                               //Extractor Cnv FROM CNV1
                           ELSIF (#Destination_Location.Device_Type = 12 AND #Source_Location.Device_Type = 10 AND
                               NOT "Control_DB".ECnv_Sys[#Id].Cnv_Occupied AND
                               "Control_DB".LCnv_Sys[#Id].Cnv_Level[#Destination_Location.Level].Cnv1.Cnv_Occupied)
                           THEN //FROM ECONVEYOR TO CNV1 OR CNV2
                               "Control_DB".ECnv_Sys[#Id].Instruction.Task_ID := INT_TO_UINT("Control_DB".WCS_OPC_Control[#Id].Task_ID);
                               "Control_DB".ECnv_Sys[#Id].Instruction.Task_Metadata := "Control_DB".WCS_OPC_Control[#Id].Task_Metadata;
                               "Control_DB".ECnv_Sys[#Id].Current_Task_Type := INT_TO_UINT("Control_DB".WCS_OPC_Control[#Id].Task_Type);
                               "Control_DB".ECnv_Sys[#Id].Instruction.Transfer_From_ID := "Control_DB".WCS_OPC_Control[#Id].Source_Location;
                               "Control_DB".ECnv_Sys[#Id].Instruction.Transfer_To_ID := "Control_DB".WCS_OPC_Control[#Id].Destination_Location;
                               IF "Control_DB".WCS_OPC_Control[#Id].Pallet_Type = 'E' AND "Control_DB".WCS_OPC_Control[#Id].Pallet_Alignment = 'L' THEN
                                   "Control_DB".ECnv_Sys[#Id].Instruction.Pallet_Type := 3;
                               ELSIF "Control_DB".WCS_OPC_Control[#Id].Pallet_Type = 'E' AND "Control_DB".WCS_OPC_Control[#Id].Pallet_Alignment = 'R' THEN
                                   "Control_DB".ECnv_Sys[#Id].Instruction.Pallet_Type := 2;
                               ELSIF "Control_DB".WCS_OPC_Control[#Id].Pallet_Type = 'E' AND "Control_DB".WCS_OPC_Control[#Id].Pallet_Alignment = 'C' THEN
                                   "Control_DB".ECnv_Sys[#Id].Instruction.Pallet_Type := 4;
                               ELSIF "Control_DB".WCS_OPC_Control[#Id].Pallet_Type = 'C' THEN
                                   "Control_DB".ECnv_Sys[#Id].Instruction.Pallet_Type := 1;
                               END_IF;

                               //Enable the conveyor and start the transfer
                               "Control_DB".ECnv_Sys[#Id].Instruction.Start_Transfer := TRUE;
                               #State_CNV := 105;

                               //Extractor Cnv FROM CNV2
                           ELSIF (#Destination_Location.Device_Type = 12 AND #Source_Location.Device_Type = 11 AND
                               NOT "Control_DB".ECnv_Sys[#Id].Cnv_Occupied AND
                               "Control_DB".LCnv_Sys[#Id].Cnv_Level[#Destination_Location.Level].Cnv2.Cnv_Occupied)
                           THEN //FROM ECONVEYOR TO CNV1 OR CNV2
                               "Control_DB".ECnv_Sys[#Id].Instruction.Task_ID := INT_TO_UINT("Control_DB".WCS_OPC_Control[#Id].Task_ID);
                               "Control_DB".ECnv_Sys[#Id].Instruction.Task_Metadata := "Control_DB".WCS_OPC_Control[#Id].Task_Metadata;
                               "Control_DB".ECnv_Sys[#Id].Current_Task_Type := INT_TO_UINT("Control_DB".WCS_OPC_Control[#Id].Task_Type);
                               "Control_DB".ECnv_Sys[#Id].Instruction.Transfer_From_ID := "Control_DB".WCS_OPC_Control[#Id].Source_Location;
                               "Control_DB".ECnv_Sys[#Id].Instruction.Transfer_To_ID := "Control_DB".WCS_OPC_Control[#Id].Destination_Location;
                               IF "Control_DB".WCS_OPC_Control[#Id].Pallet_Type = 'E' AND "Control_DB".WCS_OPC_Control[#Id].Pallet_Alignment = 'L' THEN
                                   "Control_DB".ECnv_Sys[#Id].Instruction.Pallet_Type := 3;
                               ELSIF "Control_DB".WCS_OPC_Control[#Id].Pallet_Type = 'E' AND "Control_DB".WCS_OPC_Control[#Id].Pallet_Alignment = 'R' THEN
                                   "Control_DB".ECnv_Sys[#Id].Instruction.Pallet_Type := 2;
                               ELSIF "Control_DB".WCS_OPC_Control[#Id].Pallet_Type = 'E' AND "Control_DB".WCS_OPC_Control[#Id].Pallet_Alignment = 'C' THEN
                                   "Control_DB".ECnv_Sys[#Id].Instruction.Pallet_Type := 4;
                               ELSIF "Control_DB".WCS_OPC_Control[#Id].Pallet_Type = 'C' THEN
                                   "Control_DB".ECnv_Sys[#Id].Instruction.Pallet_Type := 1;
                               END_IF;

                               //Enable the conveyor and start the transfer
                               "Control_DB".ECnv_Sys[#Id].Instruction.Start_Transfer := TRUE;
                               #State_CNV := 105;

                               //Just alignment CNV 1
                           ELSIF (#Destination_Location.Device_Type = #Source_Location.Device_Type AND
                               "Control_DB".LCnv_Sys[#Id].Cnv_Level[#Destination_Location.Level].Cnv1.Cnv_Occupied) AND
                               "Control_DB".VTD_Sys[#Id].Current_Level =  "Settings_DB".LCnv_Sys[#Id].Cnv_Level[#Destination_Location.Level].Cnv1.Cnv_Level
                           THEN
                               "Control_DB".LCnv_Sys[#Id].Cnv_Level[#Destination_Location.Level].Cnv1.Instruction.Task_ID := INT_TO_UINT("Control_DB".WCS_OPC_Control[#Id].Task_ID);
                               "Control_DB".LCnv_Sys[#Id].Cnv_Level[#Destination_Location.Level].Cnv1.Instruction.Task_Metadata := "Control_DB".WCS_OPC_Control[#Id].Task_Metadata;
                               "Control_DB".LCnv_Sys[#Id].Cnv_Level[#Destination_Location.Level].Cnv1.Current_Task_Type := INT_TO_UINT("Control_DB".WCS_OPC_Control[#Id].Task_Type);
                               "Control_DB".LCnv_Sys[#Id].Cnv_Level[#Destination_Location.Level].Cnv1.Instruction.Transfer_From_ID := "Control_DB".WCS_OPC_Control[#Id].Source_Location;
                               "Control_DB".LCnv_Sys[#Id].Cnv_Level[#Destination_Location.Level].Cnv1.Instruction.Transfer_To_ID := "Control_DB".WCS_OPC_Control[#Id].Destination_Location;
                               IF "Control_DB".WCS_OPC_Control[#Id].Pallet_Type = 'E' AND "Control_DB".WCS_OPC_Control[#Id].Pallet_Alignment = 'L' THEN
                                   "Control_DB".LCnv_Sys[#Id].Cnv_Level[#Destination_Location.Level].Cnv1.Instruction.Pallet_Type := 3;
                               ELSIF "Control_DB".WCS_OPC_Control[#Id].Pallet_Type = 'E' AND "Control_DB".WCS_OPC_Control[#Id].Pallet_Alignment = 'R' THEN
                                   "Control_DB".LCnv_Sys[#Id].Cnv_Level[#Destination_Location.Level].Cnv1.Instruction.Pallet_Type := 2;
                               END_IF;

                               //Enable the conveyor and start the transfer
                               "Control_DB".LCnv_Sys[#Id].Cnv_Level[#Destination_Location.Level].Cnv1.Instruction.Pallet_Allignment := TRUE;
                               #State_CNV := 112;

                               //Just alignment CNV 2
                           ELSIF (#Destination_Location.Device_Type = #Source_Location.Device_Type AND
                               "Control_DB".LCnv_Sys[#Id].Cnv_Level[#Destination_Location.Level].Cnv2.Cnv_Occupied) AND
                               "Control_DB".VTD_Sys[#Id].Current_Level =  "Settings_DB".LCnv_Sys[#Id].Cnv_Level[#Destination_Location.Level].Cnv2.Cnv_Level
                           THEN
                               "Control_DB".LCnv_Sys[#Id].Cnv_Level[#Destination_Location.Level].Cnv2.Instruction.Task_ID := INT_TO_UINT("Control_DB".WCS_OPC_Control[#Id].Task_ID);
                               "Control_DB".LCnv_Sys[#Id].Cnv_Level[#Destination_Location.Level].Cnv2.Instruction.Task_Metadata := "Control_DB".WCS_OPC_Control[#Id].Task_Metadata;
                               "Control_DB".LCnv_Sys[#Id].Cnv_Level[#Destination_Location.Level].Cnv2.Current_Task_Type := INT_TO_UINT("Control_DB".WCS_OPC_Control[#Id].Task_Type);
                               "Control_DB".LCnv_Sys[#Id].Cnv_Level[#Destination_Location.Level].Cnv2.Instruction.Transfer_From_ID := "Control_DB".WCS_OPC_Control[#Id].Source_Location;
                               "Control_DB".LCnv_Sys[#Id].Cnv_Level[#Destination_Location.Level].Cnv2.Instruction.Transfer_To_ID := "Control_DB".WCS_OPC_Control[#Id].Destination_Location;
                               IF "Control_DB".WCS_OPC_Control[#Id].Pallet_Type = 'E' AND "Control_DB".WCS_OPC_Control[#Id].Pallet_Alignment = 'L' THEN
                                   "Control_DB".LCnv_Sys[#Id].Cnv_Level[#Destination_Location.Level].Cnv2.Instruction.Pallet_Type := 3;
                               ELSIF "Control_DB".WCS_OPC_Control[#Id].Pallet_Type = 'E' AND "Control_DB".WCS_OPC_Control[#Id].Pallet_Alignment = 'R' THEN
                                   "Control_DB".LCnv_Sys[#Id].Cnv_Level[#Destination_Location.Level].Cnv2.Instruction.Pallet_Type := 2;
                               END_IF;

                               //Enable the conveyor and start the transfer
                               "Control_DB".LCnv_Sys[#Id].Cnv_Level[#Destination_Location.Level].Cnv2.Instruction.Pallet_Allignment := TRUE;
                               #State_CNV := 112;
                           ELSE
                               IF #Destination_Location.Device_Type = 10 AND "Control_DB".LCnv_Sys[#Id].Cnv_Level[#Destination_Location.Level].Cnv1.Cnv_Occupied THEN
                                   //Conveyor It's occupied. Check the sensors on the extractor or buffer, or verify if the pallet is misaligned.
                                   "Control_DB".LCnv_Sys[#Id].Cnv_Level[#Destination_Location.Level].Cnv1.Cnv_Errors.Error_Word_1.%X1 := TRUE;

                               ELSIF #Destination_Location.Device_Type = 10 AND "Control_DB".LCnv_Sys[#Id].Cnv_Level[#Destination_Location.Level].Cnv1.Inputs.Shuttle_High THEN
                                   //The shuttle is LID high
                                   "Control_DB".LCnv_Sys[#Id].Cnv_Level[#Destination_Location.Level].Cnv1.Cnv_Errors.Error_Word_1.%X2 := TRUE;

                               ELSIF #Destination_Location.Device_Type = 11 AND "Control_DB".LCnv_Sys[#Id].Cnv_Level[#Destination_Location.Level].Cnv2.Cnv_Occupied THEN
                                   //Conveyor It's occupied. Check the sensors on the extractor or buffer, or verify if the pallet is misaligned.
                                   "Control_DB".LCnv_Sys[#Id].Cnv_Level[#Destination_Location.Level].Cnv2.Cnv_Errors.Error_Word_1.%X1 := TRUE;

                               ELSIF #Destination_Location.Device_Type = 11 AND "Control_DB".LCnv_Sys[#Id].Cnv_Level[#Destination_Location.Level].Cnv2.Inputs.Shuttle_High THEN
                                   // The shuttle is LID high
                                   "Control_DB".LCnv_Sys[#Id].Cnv_Level[#Destination_Location.Level].Cnv2.Cnv_Errors.Error_Word_1.%X2 := TRUE;

                               ELSIF #Destination_Location.Device_Type = 12 THEN
                                   "Control_DB".ECnv_Sys[#Id].Cnv_Errors.Error_Word_1.%X1 := TRUE;
                               END_IF;

                               #State_CNV := 400; //ERROR
                           END_IF;
                       END_IF;

                   105:  //Set the source conveyor variables

                       //Assign task to sending conveyor
                       IF #Source_Location.Level >= "Settings_DB".VTD_Sys[#Id].Lowest_Level AND #Source_Location.Level <= "Settings_DB".VTD_Sys[#Id].Highest_Level THEN
                           //Cnv1
                           IF #Source_Location.Device_Type = 10 AND NOT "Control_DB".ECnv_Sys[#Id].Cnv_Occupied AND
                               "Control_DB".LCnv_Sys[#Id].Cnv_Level[#Source_Location.Level].Cnv1.Cnv_Occupied
                           THEN //FROM CONV1 TO ECONVEYOR
                               "Control_DB".LCnv_Sys[#Id].Cnv_Level[#Source_Location.Level].Cnv1.Instruction.Task_ID := INT_TO_UINT("Control_DB".WCS_OPC_Control[#Id].Task_ID);
                               "Control_DB".LCnv_Sys[#Id].Cnv_Level[#Source_Location.Level].Cnv1.Instruction.Task_Metadata := "Control_DB".WCS_OPC_Control[#Id].Task_Metadata;
                               "Control_DB".LCnv_Sys[#Id].Cnv_Level[#Source_Location.Level].Cnv1.Current_Task_Type := INT_TO_UINT("Control_DB".WCS_OPC_Control[#Id].Task_Type);
                               "Control_DB".LCnv_Sys[#Id].Cnv_Level[#Source_Location.Level].Cnv1.Instruction.Transfer_To_ID := "Control_DB".WCS_OPC_Control[#Id].Destination_Location;
                               "Control_DB".LCnv_Sys[#Id].Cnv_Level[#Source_Location.Level].Cnv1.Instruction.Transfer_From_ID := "Control_DB".WCS_OPC_Control[#Id].Source_Location;

                               //Enable the conveyor and start the transfer
                               "Control_DB".LCnv_Sys[#Id].Cnv_Level[#Source_Location.Level].Cnv1.Instruction.Start_Transfer := TRUE;
                               #State_CNV := 110;

                               //Cnv2
                           ELSIF (#Source_Location.Device_Type = 11 AND NOT "Control_DB".ECnv_Sys[#Id].Cnv_Occupied AND
                               "Control_DB".LCnv_Sys[#Id].Cnv_Level[#Source_Location.Level].Cnv2.Cnv_Occupied) OR
                               (#Source_Location.Device_Type = 11 AND #Source_Location.Level = 1 AND #Destination_Location.Device_Type = 0 AND
                               "Control_DB".LCnv_Sys[#Id].Cnv_Level[#Destination_Location.Level].Cnv2.Cnv_Occupied)
                           THEN //FROM CONV1 TO ECONVEYOR
                               "Control_DB".LCnv_Sys[#Id].Cnv_Level[#Source_Location.Level].Cnv2.Instruction.Task_ID := INT_TO_UINT("Control_DB".WCS_OPC_Control[#Id].Task_ID);
                               "Control_DB".LCnv_Sys[#Id].Cnv_Level[#Source_Location.Level].Cnv2.Instruction.Task_Metadata := "Control_DB".WCS_OPC_Control[#Id].Task_Metadata;
                               "Control_DB".LCnv_Sys[#Id].Cnv_Level[#Source_Location.Level].Cnv2.Current_Task_Type := INT_TO_UINT("Control_DB".WCS_OPC_Control[#Id].Task_Type);
                               "Control_DB".LCnv_Sys[#Id].Cnv_Level[#Source_Location.Level].Cnv2.Instruction.Transfer_To_ID := "Control_DB".WCS_OPC_Control[#Id].Destination_Location;
                               "Control_DB".LCnv_Sys[#Id].Cnv_Level[#Source_Location.Level].Cnv2.Instruction.Transfer_From_ID := "Control_DB".WCS_OPC_Control[#Id].Source_Location;

                               //Enable the conveyor and start the transfer
                               "Control_DB".LCnv_Sys[#Id].Cnv_Level[#Source_Location.Level].Cnv2.Instruction.Start_Transfer := TRUE;
                               #State_CNV := 110;

                               //Extractor Cnv TO CNV 1
                           ELSIF (#Source_Location.Device_Type = 12 AND #Destination_Location.Device_Type = 10 AND "Control_DB".ECnv_Sys[#Id].Cnv_Occupied AND
                               NOT "Control_DB".LCnv_Sys[#Id].Cnv_Level[#Source_Location.Level].Cnv1.Cnv_Occupied)
                           THEN //FROM ECONVEYOR TO CNV1
                               "Control_DB".ECnv_Sys[#Id].Instruction.Task_ID := INT_TO_UINT("Control_DB".WCS_OPC_Control[#Id].Task_ID);
                               "Control_DB".ECnv_Sys[#Id].Instruction.Task_Metadata := "Control_DB".WCS_OPC_Control[#Id].Task_Metadata;
                               "Control_DB".ECnv_Sys[#Id].Current_Task_Type := INT_TO_UINT("Control_DB".WCS_OPC_Control[#Id].Task_Type);
                               "Control_DB".ECnv_Sys[#Id].Instruction.Transfer_To_ID := "Control_DB".WCS_OPC_Control[#Id].Destination_Location;
                               "Control_DB".ECnv_Sys[#Id].Instruction.Transfer_From_ID := "Control_DB".WCS_OPC_Control[#Id].Source_Location;

                               //Enable the conveyor and start the transfer
                               "Control_DB".ECnv_Sys[#Id].Instruction.Start_Transfer := TRUE;
                               #State_CNV := 110;

                               //Extractor Cnv TO CNV 2
                           ELSIF (#Source_Location.Device_Type = 12 AND #Destination_Location.Device_Type = 11 AND "Control_DB".ECnv_Sys[#Id].Cnv_Occupied AND
                               NOT "Control_DB".LCnv_Sys[#Id].Cnv_Level[#Source_Location.Level].Cnv2.Cnv_Occupied)
                           THEN //FROM ECONVEYOR TO CNV2
                               "Control_DB".ECnv_Sys[#Id].Instruction.Task_ID := INT_TO_UINT("Control_DB".WCS_OPC_Control[#Id].Task_ID);
                               "Control_DB".ECnv_Sys[#Id].Instruction.Task_Metadata := "Control_DB".WCS_OPC_Control[#Id].Task_Metadata;
                               "Control_DB".ECnv_Sys[#Id].Current_Task_Type := INT_TO_UINT("Control_DB".WCS_OPC_Control[#Id].Task_Type);
                               "Control_DB".ECnv_Sys[#Id].Instruction.Transfer_To_ID := "Control_DB".WCS_OPC_Control[#Id].Destination_Location;
                               "Control_DB".ECnv_Sys[#Id].Instruction.Transfer_From_ID := "Control_DB".WCS_OPC_Control[#Id].Source_Location;

                               //Enable the conveyor and start the transfer
                               "Control_DB".ECnv_Sys[#Id].Instruction.Start_Transfer := TRUE;
                               #State_CNV := 110;
                           ELSE
                               #State_CNV := 400; //ERROR
                           END_IF;
                       ELSE
                           #State_CNV := 400;
                       END_IF;

                   110: //Start the transfer
                       "Control_DB".WCS_OPC_Control[#Id].SM_State := "Control_DB".ECnv_Sys[#Id].SM_State;

                       IF "Control_DB".ECnv_Sys[#Id].Enabled AND "Control_DB".ECnv_Sys[#Id].Running
                       THEN
                           "Control_DB".ECnv_Sys[#Id].Instruction.Start_Transfer := FALSE;
                           IF (#Source_Location.Device_Type = 12 AND #Destination_Location.Device_Type = 10) OR
                               (#Source_Location.Device_Type = 10 AND #Destination_Location.Device_Type = 12) AND
                               "Control_DB".LCnv_Sys[#Id].Cnv_Level["Control_DB".VTD_Sys[#Id].Current_Level].Cnv1.Running
                           THEN
                               "Control_DB".LCnv_Sys[#Id].Cnv_Level["Control_DB".VTD_Sys[#Id].Current_Level].Cnv1.Instruction.Start_Transfer := FALSE;
                               #State_CNV := 115;
                           ELSIF (#Source_Location.Device_Type = 12 AND #Destination_Location.Device_Type = 11) OR
                               (#Source_Location.Device_Type = 11 AND #Destination_Location.Device_Type = 12) AND
                               "Control_DB".LCnv_Sys[#Id].Cnv_Level["Control_DB".VTD_Sys[#Id].Current_Level].Cnv2.Running
                           THEN
                               "Control_DB".LCnv_Sys[#Id].Cnv_Level["Control_DB".VTD_Sys[#Id].Current_Level].Cnv2.Instruction.Start_Transfer := FALSE;
                               #State_CNV := 115;
                           END_IF;
                           "Control_DB".WCS_OPC_Control[#Id].Movement_Ready := TRUE;
                       END_IF;

                   112: //Start the transfer
                       IF "Control_DB".LCnv_Sys[#Id].Cnv_Level[#Destination_Location.Level].Cnv1.Enabled AND "Control_DB".LCnv_Sys[#Id].Cnv_Level[#Destination_Location.Level].Cnv1.Running
                       THEN
                           "Control_DB".WCS_OPC_Control[#Id].SM_State := "Control_DB".LCnv_Sys[#Id].Cnv_Level[#Destination_Location.Level].Cnv1.SM_State;
                           "Control_DB".LCnv_Sys[#Id].Cnv_Level[#Destination_Location.Level].Cnv1.Instruction.Pallet_Allignment := FALSE;
                           "Control_DB".WCS_OPC_Control[#Id].Movement_Ready := TRUE;
                           #State_CNV := 116;
                       ELSIF "Control_DB".LCnv_Sys[#Id].Cnv_Level[#Destination_Location.Level].Cnv2.Enabled AND "Control_DB".LCnv_Sys[#Id].Cnv_Level[#Destination_Location.Level].Cnv2.Running
                       THEN
                           "Control_DB".WCS_OPC_Control[#Id].SM_State := "Control_DB".LCnv_Sys[#Id].Cnv_Level[#Destination_Location.Level].Cnv2.SM_State;
                           "Control_DB".LCnv_Sys[#Id].Cnv_Level[#Destination_Location.Level].Cnv2.Instruction.Pallet_Allignment := FALSE;
                           "Control_DB".WCS_OPC_Control[#Id].Movement_Ready := TRUE;
                           #State_CNV := 116;
                       END_IF;



                   115: //Wait for the transfer to complete
                       "Control_DB".WCS_OPC_Control[#Id].SM_State := "Control_DB".ECnv_Sys[#Id].SM_State;
                       IF (#Source_Location.Device_Type = 12 AND #Destination_Location.Device_Type = 10) OR
                           (#Source_Location.Device_Type = 10 AND #Destination_Location.Device_Type = 12) THEN
                           IF "Control_DB".ECnv_Sys[#Id].Done AND "Control_DB".LCnv_Sys[#Id].Cnv_Level[#Destination_Location.Level].Cnv1.Done THEN
                               #State_CNV := 118;
                           END_IF;
                       ELSIF (#Source_Location.Device_Type = 12 AND #Destination_Location.Device_Type = 11) OR
                           (#Source_Location.Device_Type = 11 AND #Destination_Location.Device_Type = 12) THEN
                           IF "Control_DB".ECnv_Sys[#Id].Done AND "Control_DB".LCnv_Sys[#Id].Cnv_Level[#Destination_Location.Level].Cnv2.Done THEN
                               #State_CNV := 118;
                           END_IF;
                       END_IF;

                   116: //Wait for the ALIGNMENT to complete
                           IF "Control_DB".LCnv_Sys[#Id].Cnv_Level[#Destination_Location.Level].Cnv1.Done THEN
                               #State_CNV := 118;
                           END_IF;
                           IF "Control_DB".LCnv_Sys[#Id].Cnv_Level[#Destination_Location.Level].Cnv2.Done THEN
                               #State_CNV := 118;
                           END_IF;

                   118: //Wait for XXs for report done
                       #T_Wait_Report_Done.TON(IN := TRUE,
                                              PT := T#500mS);
                      IF #T_Wait_Report_Done.Q THEN
                           "Control_DB".WCS_OPC_Control[#Id].Movement_Request_Complete := TRUE;
                           #State_CNV := 120;
                       END_IF;

                   120: //Wait for the ACK before we go back to Idle
                       "Control_DB".WCS_OPC_Control[#Id].SM_State := "Control_DB".ECnv_Sys[#Id].SM_State;
                       IF "Control_DB".WCS_OPC_Control[#Id].Movement_Request_Complete_Ack THEN
                           #State_CNV := 250;
                       END_IF;

                   250: //Reset all variable and return to idle
                       "Control_DB".ECnv_Sys[#Id].Instruction.Reset := FALSE;
                       "Control_DB".ECnv_Sys[#Id].Instruction.Start_Transfer := FALSE;
                       "Control_DB".ECnv_Sys[#Id].Instruction.Task_ID := 0;
                       "Control_DB".ECnv_Sys[#Id].Instruction.Task_Metadata := '';
                       "Control_DB".ECnv_Sys[#Id].Current_Task_Type := 0;
                       "Control_DB".ECnv_Sys[#Id].Instruction.Transfer_From_ID := 0;
                       "Control_DB".ECnv_Sys[#Id].Instruction.Transfer_To_ID := 0;
                       IF #Destination_Location.Device_Type = 10 THEN
                           "Control_DB".LCnv_Sys[#Id].Cnv_Level[#Destination_Location.Level].Cnv1.Instruction.Reset := FALSE;
                           "Control_DB".LCnv_Sys[#Id].Cnv_Level[#Destination_Location.Level].Cnv1.Instruction.Start_Transfer := FALSE;
                           "Control_DB".LCnv_Sys[#Id].Cnv_Level[#Destination_Location.Level].Cnv1.Instruction.Task_ID := 0;
                           "Control_DB".LCnv_Sys[#Id].Cnv_Level[#Destination_Location.Level].Cnv1.Instruction.Task_Metadata := '';
                           "Control_DB".LCnv_Sys[#Id].Cnv_Level[#Destination_Location.Level].Cnv1.Current_Task_Type := 0;
                           "Control_DB".LCnv_Sys[#Id].Cnv_Level[#Destination_Location.Level].Cnv1.Instruction.Transfer_From_ID := 0;
                           "Control_DB".LCnv_Sys[#Id].Cnv_Level[#Destination_Location.Level].Cnv1.Instruction.Transfer_To_ID := 0;
                       ELSIF #Destination_Location.Device_Type = 11 THEN
                           "Control_DB".LCnv_Sys[#Id].Cnv_Level[#Destination_Location.Level].Cnv2.Instruction.Reset := FALSE;
                           "Control_DB".LCnv_Sys[#Id].Cnv_Level[#Destination_Location.Level].Cnv2.Instruction.Start_Transfer := FALSE;
                           "Control_DB".LCnv_Sys[#Id].Cnv_Level[#Destination_Location.Level].Cnv2.Instruction.Task_ID := 0;
                           "Control_DB".LCnv_Sys[#Id].Cnv_Level[#Destination_Location.Level].Cnv2.Instruction.Task_Metadata := '';
                           "Control_DB".LCnv_Sys[#Id].Cnv_Level[#Destination_Location.Level].Cnv2.Current_Task_Type := 0;
                           "Control_DB".LCnv_Sys[#Id].Cnv_Level[#Destination_Location.Level].Cnv2.Instruction.Transfer_From_ID := 0;
                           "Control_DB".LCnv_Sys[#Id].Cnv_Level[#Destination_Location.Level].Cnv2.Instruction.Transfer_To_ID := 0;
                       ELSIF #Source_Location.Device_Type = 10 THEN
                           "Control_DB".LCnv_Sys[#Id].Cnv_Level[#Source_Location.Level].Cnv1.Instruction.Reset := FALSE;
                           "Control_DB".LCnv_Sys[#Id].Cnv_Level[#Source_Location.Level].Cnv1.Instruction.Start_Transfer := FALSE;
                           "Control_DB".LCnv_Sys[#Id].Cnv_Level[#Source_Location.Level].Cnv1.Instruction.Task_ID := 0;
                           "Control_DB".LCnv_Sys[#Id].Cnv_Level[#Source_Location.Level].Cnv1.Instruction.Task_Metadata := '';
                           "Control_DB".LCnv_Sys[#Id].Cnv_Level[#Source_Location.Level].Cnv1.Current_Task_Type := 0;
                           "Control_DB".LCnv_Sys[#Id].Cnv_Level[#Source_Location.Level].Cnv1.Instruction.Transfer_From_ID := 0;
                           "Control_DB".LCnv_Sys[#Id].Cnv_Level[#Source_Location.Level].Cnv1.Instruction.Transfer_To_ID := 0;
                       ELSIF #Destination_Location.Device_Type = 11 THEN
                           "Control_DB".LCnv_Sys[#Id].Cnv_Level[#Source_Location.Level].Cnv2.Instruction.Reset := FALSE;
                           "Control_DB".LCnv_Sys[#Id].Cnv_Level[#Source_Location.Level].Cnv2.Instruction.Start_Transfer := FALSE;
                           "Control_DB".LCnv_Sys[#Id].Cnv_Level[#Source_Location.Level].Cnv2.Instruction.Task_ID := 0;
                           "Control_DB".LCnv_Sys[#Id].Cnv_Level[#Source_Location.Level].Cnv2.Instruction.Task_Metadata := '';
                           "Control_DB".LCnv_Sys[#Id].Cnv_Level[#Source_Location.Level].Cnv2.Current_Task_Type := 0;
                           "Control_DB".LCnv_Sys[#Id].Cnv_Level[#Source_Location.Level].Cnv2.Instruction.Transfer_From_ID := 0;
                           "Control_DB".LCnv_Sys[#Id].Cnv_Level[#Source_Location.Level].Cnv2.Instruction.Transfer_To_ID := 0;
                       END_IF;

                       // IF (#State_VTD = 0 OR #State_VTD = 250) AND
                       //     (#State_Shuttle = 0 OR #State_Shuttle = 250) THEN
                           //Reset the OPC control variables
                           "Control_DB".WCS_OPC_Control[#Id].SM_State := 0;
                           "Control_DB".WCS_OPC_Control[#Id].Movement_Ready := FALSE;
                           "Control_DB".WCS_OPC_Control[#Id].Movement_Request_Complete := FALSE;
                           "Control_DB".WCS_OPC_Control[#Id].Movement_Request_Complete_Ack := FALSE;
                           "Control_DB".WCS_OPC_Control[#Id].Task_Metadata := '';
                           #T_Wait_Report_Done.TON(IN := FALSE,
                                                  PT := T#0S);

                           #State_CNV := 0;
                       // END_IF;

                       400:// Error state
                           #Error_ID.%X8 := TRUE;
                           IF "Reset_All" OR #HMI_Reset THEN
                               #Error_ID.%X3 := FALSE;
                               #Error_ID.%X4 := FALSE;
                               #Error_ID.%X8 := FALSE;
                               #State_CNV := 250;
                       END_IF;
               END_CASE;
           END_REGION ;
       END_REGION

   ELSIF #All_In_Automatic AND NOT #OPC_Enable THEN
       //Reset all variable and return to idle

       //Reset the OPC control variables
       "Control_DB".WCS_OPC_Control[#Id].SM_State := 0;
       "Control_DB".WCS_OPC_Control[#Id].Movement_Ready := FALSE;
       "Control_DB".WCS_OPC_Control[#Id].Movement_Request_Complete := FALSE;

       // Reset Order table VTD variables
       "Control_DB".WCS_OPC_Control[#Id].Task_Type := 0;
       "Control_DB".WCS_OPC_Control[#Id].Pallet_Type := 'C';
       "Control_DB".WCS_OPC_Control[#Id].Task_ID := 0;
       "Control_DB".WCS_OPC_Control[#Id].Task_Metadata := '';
       "Control_DB".WCS_OPC_Control[#Id].Source_Location := 0;
       "Control_DB".WCS_OPC_Control[#Id].Destination_Location := 0;
       #Destination_Location.Level := 0;
       #Source_Location.Level := 0;
       "Control_DB".WCS_OPC_Control[#Id].Shuttle_ID := 0;
       "Control_DB".WCS_OPC_Control[#Id].Shuttle_Loaded := FALSE;

       //Reset VTD variables
       "Control_DB".VTD_Sys[#Id].Instruction.Reset := FALSE;
       "Control_DB".VTD_Sys[#Id].Instruction.Pallet_Type := 0;
       "Control_DB".VTD_Sys[#Id].Instruction.Task_ID := 0;
       "Control_DB".VTD_Sys[#Id].Instruction.Task_Metadata := '';//
       "Control_DB".ECnv_Sys[#Id].Current_Task_Type := 0;
       "Control_DB".VTD_Sys[#Id].Instruction.Move_To_Level := 99;
       "Control_DB".VTD_Sys[#Id].Current_Task_Type := 0;

       //Reset Shuttle interlock
       "Control_DB".VTD_Sys[#Id].Shuttle_Interlock.Interlock_Request := FALSE;
       "Control_DB".VTD_Sys[#Id].Shuttle_Interlock.Shuttle_Start_Location := 0;
       "Control_DB".VTD_Sys[#Id].Shuttle_Interlock.Shuttle_Target_Location := 0;
       "Control_DB".VTD_Sys[#Id].Shuttle_Interlock.Shuttle_Loaded := 0;
       "Control_DB".VTD_Sys[#Id].Shuttle_Interlock.Shuttle_ID := 0;
       "Control_DB".VTD_Sys[#Id].Shuttle_Interlock.Shuttle_Interlock_Task_ID := 0;
       "Control_DB".VTD_Sys[#Id].Shuttle_Interlock.Shuttle_Interlock_Task_Metadata := '';//

       //Reset conveyor variables
       "Control_DB".ECnv_Sys[#Id].Instruction.Reset := FALSE;
       // "Control_DB".ECnv_Control.Instruction.Enable := FALSE;
       "Control_DB".ECnv_Sys[#Id].Instruction.Start_Transfer := FALSE;
       "Control_DB".ECnv_Sys[#Id].Instruction.Task_ID := 0;
       "Control_DB".ECnv_Sys[#Id].Instruction.Task_Metadata := '';//
       "Control_DB".ECnv_Sys[#Id].Instruction.Transfer_From_ID := 0;
       "Control_DB".ECnv_Sys[#Id].Instruction.Transfer_To_ID := 0;

       FOR #i := "Settings_DB".VTD_Sys[#Id].Lowest_Level TO "Settings_DB".VTD_Sys[#Id].Highest_Level DO
           "Control_DB".LCnv_Sys[#Id].Cnv_Level[#i].Cnv1.Instruction.Reset := FALSE;
           "Control_DB".LCnv_Sys[#Id].Cnv_Level[#i].Cnv1.Instruction.Start_Transfer := FALSE;
           "Control_DB".LCnv_Sys[#Id].Cnv_Level[#i].Cnv1.Instruction.Task_ID := 0;
           "Control_DB".LCnv_Sys[#Id].Cnv_Level[#i].Cnv1.Instruction.Task_Metadata := '';
           "Control_DB".LCnv_Sys[#Id].Cnv_Level[#i].Cnv1.Current_Task_Type := 0;
           "Control_DB".LCnv_Sys[#Id].Cnv_Level[#i].Cnv1.Instruction.Transfer_From_ID := 0;
           "Control_DB".LCnv_Sys[#Id].Cnv_Level[#i].Cnv1.Instruction.Transfer_To_ID := 0;

           "Control_DB".LCnv_Sys[#Id].Cnv_Level[#i].Cnv2.Instruction.Reset := FALSE;
           "Control_DB".LCnv_Sys[#Id].Cnv_Level[#i].Cnv2.Instruction.Start_Transfer := FALSE;
           "Control_DB".LCnv_Sys[#Id].Cnv_Level[#i].Cnv2.Instruction.Task_ID := 0;
           "Control_DB".LCnv_Sys[#Id].Cnv_Level[#i].Cnv2.Instruction.Task_Metadata := '';
           "Control_DB".LCnv_Sys[#Id].Cnv_Level[#i].Cnv2.Current_Task_Type := 0;
           "Control_DB".LCnv_Sys[#Id].Cnv_Level[#i].Cnv2.Instruction.Transfer_From_ID := 0;
           "Control_DB".LCnv_Sys[#Id].Cnv_Level[#i].Cnv2.Instruction.Transfer_To_ID := 0;
       END_FOR;
   END_IF;

   REGION Clear order table
       IF #Clear_OrderTable THEN
           #State_Main := 0;
           #State_VTD := 250;
           #State_Shuttle := 250;
           #State_CNV := 250;
           "Control_DB".WCS_OPC_Control[#Id].Task_Data_Available := 0;
       END_IF;
   END_REGION

   REGION SHUTTLES POSITION
       FOR #f := 1 TO "Settings_DB".System.Shuttle_Count DO
           "Control_DB".Shuttles_Position[#f].x := "Shuttle_MQTT_DB".Shuttle_MQTT[#f].Message.Shuttle_Status.Position_X;
           "Control_DB".Shuttles_Position[#f].y := "Shuttle_MQTT_DB".Shuttle_MQTT[#f].Message.Shuttle_Status.Position_Y;
       END_FOR;
   END_REGION

   REGION SM STATE MAESTRO
       // Statement section - Send the State machine to Maestro "Emulating" openTCS states
       // 
       // // "Control_DB".WMS_OPC_UA.SM_State_Maestro; // State to send Devices to Maestro
       //  IF #State_VTD = 0 THEN

       //      "Control_DB"."Order Table"[#Id].SM_State_Maestro := 0;//"LIMBO" condition 

       //  ELSIF "Control_DB"."Order Table"[#Id].SM_State = 10 THEN
       //      ;
       //      // "Control_DB".WMS_OPC_UA.SM_State_Maestro := 1;//RAW conidtion => Maestro will write this condition

       //      //////////////////////////////////////////////////////////////////////////////////////////////////////////////////////      
       //      // QUEUED ANY DEVICE    
       //  // ELSIF "Control_DB".WMS_OPC_UA.Task_Data_Available AND #State >= 10 AND #State <= 20 THEN
       //  ELSIF "Control_DB"."Order Table"[#Id].Task_Data_Available AND NOT "Control_DB"."Order Table"[#Id].Movement_Ready AND "Control_DB"."Order Table"[#Id].SM_State_Maestro = 1 THEN
       //      "Control_DB"."Order Table"[#Id].SM_State_Maestro := 2;//QUEUED condition =>ANY device (Conveyor, VTD OR Shuttle)  

       //      //////////////////////////////////////////////////////////////////////////////////////////////////////////////////////       
       //      // Any Device RUNNING on the system (VTD - Conveyor Transfer - Shuttle Transfer) 
       //  ELSIF ("Control_DB"."Order Table"[#Id].Task_Type = 4 OR "Control_DB"."Order Table"[#Id].Task_Type = 5
       //      OR "Control_DB"."Order Table"[#Id].Task_Type = 1 OR "Control_DB"."Order Table"[#Id].Task_Type = 2 OR "Control_DB"."Order Table"[#Id].Task_Type = 3)
       //      AND "Control_DB"."Order Table"[#Id].Movement_Ready AND NOT "Control_DB"."Order Table"[#Id].Movement_Request_Complete THEN

       //      "Control_DB"."Order Table"[#Id].SM_State_Maestro := 3;//RUNNING condition

       //      // Any Device DONE on the system (VTD - Coneveyor Transfer - Shuttle Transfer) 
       //  ELSIF ("Control_DB"."Order Table"[#Id].Task_Type = 4 OR "Control_DB"."Order Table"[#Id].Task_Type = 5
       //      OR "Control_DB"."Order Table"[#Id].Task_Type = 1 OR "Control_DB"."Order Table"[#Id].Task_Type = 2 OR "Control_DB"."Order Table"[#Id].Task_Type = 3)
       //      AND (*"Control_DB".WMS_OPC_UA.Movement_Request_Complete AND "Control_DB".WMS_OPC_UA.Movement_Ready*)#State_VTD = 120 OR #State_VTD = 45 OR #State_VTD = 90 THEN

       //      "Control_DB"."Order Table"[#Id].SM_State_Maestro := 4;//DONE condition

       //      // Any Device ERRORS on the system (VTD - Coneveyor Transfer - Shuttle Transfer)  
       //  ELSIF ("Control_DB"."Order Table"[#Id].Task_Type = 4 OR "Control_DB"."Order Table"[#Id].Task_Type = 5
       //      OR "Control_DB"."Order Table"[#Id].Task_Type = 1 OR "Control_DB"."Order Table"[#Id].Task_Type = 2 OR "Control_DB"."Order Table"[#Id].Task_Type = 3)
       //      AND "Control_DB"."Order Table"[#Id].SM_State = 400 THEN

       //      "Control_DB"."Order Table"[#Id].SM_State_Maestro := 5;//ERROR condition => Conveyors   
       //  END_IF;
       //      /////////////////////////////////////////////////////////////////////////////////////////////        



       // "Control_DB".WMS_OPC_UA.SM_State_Maestro; // State to send Devices to Maestro
       // IF #State_Main = 0 THEN
       //     ;
       //     //"System_DB_VTD".OrderTable[1].OPC_Control.SM_State_Maestro := 0;//"LIMBO" condition 

       // ELSIF "Control_DB".WCS_OPC_Control[#Id].SM_State = 10 THEN
       //     ;
       //     // "Control_DB".WMS_OPC_UA.SM_State_Maestro := 1;//RAW conidtion => Maestro will write this condition

       //     //////////////////////////////////////////////////////////////////////////////////////////////////////////////////////      
       //     // QUEUED ANY DEVICE    
       //     // ELSIF "Control_DB".WMS_OPC_UA.Task_Data_Available AND #State >= 10 AND #State <= 20 THEN
       // ELSIF "Control_DB".WCS_OPC_Control[#Id].Task_Data_Available AND NOT "Control_DB".WCS_OPC_Control[#Id].Movement_Ready AND "System_DB_1".OrderTable[1].OPC_Control.SM_State_Maestro = 1 THEN
       //     "System_DB_1".OrderTable[1].OPC_Control.SM_State_Maestro := 2;//QUEUED condition =>ANY device (Conveyor, VTD OR Shuttle)  

       //     //////////////////////////////////////////////////////////////////////////////////////////////////////////////////////       
       //     // Any Device RUNNING on the system (VTD - Conveyor Transfer - Shuttle Transfer) 
       // ELSIF ("Control_DB".WCS_OPC_Control[#Id].Task_Type = 4 OR "Control_DB".WCS_OPC_Control[#Id].Task_Type = 5
       //     OR "Control_DB".WCS_OPC_Control[#Id].Task_Type = 1 OR "Control_DB".WCS_OPC_Control[#Id].Task_Type = 2 OR "Control_DB".WCS_OPC_Control[#Id].Task_Type = 3)
       //     AND "Control_DB".WCS_OPC_Control[#Id].Movement_Ready AND NOT "Control_DB".WCS_OPC_Control[#Id].Movement_Request_Complete THEN

       //     "System_DB_1".OrderTable[1].OPC_Control.SM_State_Maestro := 3;//RUNNING condition

       //     // Any Device DONE on the system (VTD - Coneveyor Transfer - Shuttle Transfer) 
       // ELSIF ("Control_DB".WCS_OPC_Control[#Id].Task_Type = 4 OR "Control_DB".WCS_OPC_Control[#Id].Task_Type = 5
       //     OR "Control_DB".WCS_OPC_Control[#Id].Task_Type = 1 OR "Control_DB".WCS_OPC_Control[#Id].Task_Type = 2 OR "Control_DB".WCS_OPC_Control[#Id].Task_Type = 3)
       //     AND (*"Control_DB".WMS_OPC_UA.Movement_Request_Complete AND "Control_DB".WMS_OPC_UA.Movement_Ready*)#State_Main = 120 OR #State_Main = 45 OR #State_Main = 90 THEN

       //     "System_DB_1".OrderTable[1].OPC_Control.SM_State_Maestro := 4;//DONE condition

       //     // Any Device ERRORS on the system (VTD - Coneveyor Transfer - Shuttle Transfer)  
       // ELSIF ("Control_DB".WCS_OPC_Control[#Id].Task_Type = 4 OR "Control_DB".WCS_OPC_Control[#Id].Task_Type = 5
       //     OR "Control_DB".WCS_OPC_Control[#Id].Task_Type = 1 OR "Control_DB".WCS_OPC_Control[#Id].Task_Type = 2 OR "Control_DB".WCS_OPC_Control[#Id].Task_Type = 3)
       //     AND "Control_DB".WCS_OPC_Control[#Id].SM_State = 400 THEN

       //     "System_DB_1".OrderTable[1].OPC_Control.SM_State_Maestro := 5;//ERROR condition => Conveyors   
       // END_IF;
       /////////////////////////////////////////////////////////////////////////////////////////////        


       //  //     //////////////////////////////////////////////////////////////////////////////////////////////////////////////////////       
       //  //     // Any VTD RUNNING on the system (VTD) 
       //  // ELSIF "Control_DB".WMS_OPC_UA.Task_Type = 1
       //  //     AND "Control_DB".WMS_OPC_UA.SM_State >= 35 AND "Control_DB".WMS_OPC_UA.SM_State < 100 AND #State > 20 THEN

       //  //     "Control_DB".WMS_OPC_UA.SM_State_Maestro := 3;//RUNNING condition => VTD

       //  //     // Any VTD DONE on the system (VTD) 
       //  // ELSIF "Control_DB".WMS_OPC_UA.Task_Type = 1
       //  //     AND "Control_DB".WMS_OPC_UA.SM_State = 100 AND #State > 20 THEN

       //  //     "Control_DB".WMS_OPC_UA.SM_State_Maestro := 4;//DONE condition => VTD

       //  //     // Any VTD ERRORS on the system (VTD) 
       //  // ELSIF "Control_DB".WMS_OPC_UA.Task_Type = 1
       //  //     AND "Control_DB".WMS_OPC_UA.SM_State = 400 THEN

       //  //     "Control_DB".WMS_OPC_UA.SM_State_Maestro := 5;//ERROR condition => VTD   



       //  //     //////////////////////////////////////////////////////////////////////////////////////////////////////////////////////       
       //  //     // Any Shuttle Interlock RUNNING on the system (Shuttle) 
       //  // ELSIF "Control_DB".WMS_OPC_UA.Task_Type = 2 OR "Control_DB".WMS_OPC_UA.Task_Type = 3
       //  //     AND "Control_DB".WMS_OPC_UA.SM_State >= 35 AND "Control_DB".WMS_OPC_UA.SM_State < 100 AND #State > 20 THEN

       //  //     "Control_DB".WMS_OPC_UA.SM_State_Maestro := 3;//RUNNING condition => Shuttle

       //  //     // Any Shuttle Interlock  DONE on the system (Shuttle) 
       //  // ELSIF "Control_DB".WMS_OPC_UA.Task_Type = 2 OR "Control_DB".WMS_OPC_UA.Task_Type = 3
       //  //     AND "Control_DB".WMS_OPC_UA.SM_State = 100 AND #State > 20 THEN

       //  //     "Control_DB".WMS_OPC_UA.SM_State_Maestro := 4;//DONE condition => Shuttle

       //  //     // Any Shuttle Interlock ERRORS on the system (Shuttle) 
       //  // ELSIF "Control_DB".WMS_OPC_UA.Task_Type = 2 OR "Control_DB".WMS_OPC_UA.Task_Type = 3
       //  //     AND "Control_DB".WMS_OPC_UA.SM_State = 400 THEN

       //  //     "Control_DB".WMS_OPC_UA.SM_State_Maestro := 5;//ERROR condition => Shuttle          

       //  // END_IF;


       // // "Control_DB".WMS_OPC_UA.SM_State_Maestro; // State to send Devices to Maestro
       //  IF #State_VTD = 0 THEN

       //      "Control_DB"."Order Table"[#Id].SM_State_Maestro := 0;//"LIMBO" condition 

       //  ELSIF "Control_DB"."Order Table"[#Id].SM_State = 10 THEN
       //      ;
       //      // "Control_DB".WMS_OPC_UA.SM_State_Maestro := 1;//RAW conidtion => Maestro will write this condition

       //      //////////////////////////////////////////////////////////////////////////////////////////////////////////////////////      
       //      // QUEUED ANY DEVICE    
       //  // ELSIF "Control_DB".WMS_OPC_UA.Task_Data_Available AND #State >= 10 AND #State <= 20 THEN
       //  ELSIF "Control_DB"."Order Table"[#Id].Task_Data_Available AND NOT "Control_DB"."Order Table"[#Id].Movement_Ready AND "Control_DB"."Order Table"[#Id].SM_State_Maestro = 1 THEN
       //      "Control_DB"."Order Table"[#Id].SM_State_Maestro := 2;//QUEUED condition =>ANY device (Conveyor, VTD OR Shuttle)  

       //      //////////////////////////////////////////////////////////////////////////////////////////////////////////////////////       
       //      // Any Device RUNNING on the system (VTD - Conveyor Transfer - Shuttle Transfer) 
       //  ELSIF ("Control_DB"."Order Table"[#Id].Task_Type = 4 OR "Control_DB"."Order Table"[#Id].Task_Type = 5
       //      OR "Control_DB"."Order Table"[#Id].Task_Type = 1 OR "Control_DB"."Order Table"[#Id].Task_Type = 2 OR "Control_DB"."Order Table"[#Id].Task_Type = 3)
       //      AND "Control_DB"."Order Table"[#Id].Movement_Ready AND NOT "Control_DB"."Order Table"[#Id].Movement_Request_Complete THEN

       //      "Control_DB"."Order Table"[#Id].SM_State_Maestro := 3;//RUNNING condition

       //      // Any Device DONE on the system (VTD - Coneveyor Transfer - Shuttle Transfer) 
       //  ELSIF ("Control_DB"."Order Table"[#Id].Task_Type = 4 OR "Control_DB"."Order Table"[#Id].Task_Type = 5
       //      OR "Control_DB"."Order Table"[#Id].Task_Type = 1 OR "Control_DB"."Order Table"[#Id].Task_Type = 2 OR "Control_DB"."Order Table"[#Id].Task_Type = 3)
       //      AND (*"Control_DB".WMS_OPC_UA.Movement_Request_Complete AND "Control_DB".WMS_OPC_UA.Movement_Ready*)#State_VTD = 120 OR #State_VTD = 45 OR #State_VTD = 90 THEN

       //      "Control_DB"."Order Table"[#Id].SM_State_Maestro := 4;//DONE condition

       //      // Any Device ERRORS on the system (VTD - Coneveyor Transfer - Shuttle Transfer)  
       //  ELSIF ("Control_DB"."Order Table"[#Id].Task_Type = 4 OR "Control_DB"."Order Table"[#Id].Task_Type = 5
       //      OR "Control_DB"."Order Table"[#Id].Task_Type = 1 OR "Control_DB"."Order Table"[#Id].Task_Type = 2 OR "Control_DB"."Order Table"[#Id].Task_Type = 3)
       //      AND "Control_DB"."Order Table"[#Id].SM_State = 400 THEN

       //      "Control_DB"."Order Table"[#Id].SM_State_Maestro := 5;//ERROR condition => Conveyors   
       //  END_IF;
       //      /////////////////////////////////////////////////////////////////////////////////////////////        

       //  //     //////////////////////////////////////////////////////////////////////////////////////////////////////////////////////       
       //  //     // Any VTD RUNNING on the system (VTD) 
       //  // ELSIF "Control_DB".WMS_OPC_UA.Task_Type = 1
       //  //     AND "Control_DB".WMS_OPC_UA.SM_State >= 35 AND "Control_DB".WMS_OPC_UA.SM_State < 100 AND #State > 20 THEN

       //  //     "Control_DB".WMS_OPC_UA.SM_State_Maestro := 3;//RUNNING condition => VTD

       //  //     // Any VTD DONE on the system (VTD) 
       //  // ELSIF "Control_DB".WMS_OPC_UA.Task_Type = 1
       //  //     AND "Control_DB".WMS_OPC_UA.SM_State = 100 AND #State > 20 THEN

       //  //     "Control_DB".WMS_OPC_UA.SM_State_Maestro := 4;//DONE condition => VTD

       //  //     // Any VTD ERRORS on the system (VTD) 
       //  // ELSIF "Control_DB".WMS_OPC_UA.Task_Type = 1
       //  //     AND "Control_DB".WMS_OPC_UA.SM_State = 400 THEN

       //  //     "Control_DB".WMS_OPC_UA.SM_State_Maestro := 5;//ERROR condition => VTD   



       //  //     //////////////////////////////////////////////////////////////////////////////////////////////////////////////////////       
       //  //     // Any Shuttle Interlock RUNNING on the system (Shuttle) 
       //  // ELSIF "Control_DB".WMS_OPC_UA.Task_Type = 2 OR "Control_DB".WMS_OPC_UA.Task_Type = 3
       //  //     AND "Control_DB".WMS_OPC_UA.SM_State >= 35 AND "Control_DB".WMS_OPC_UA.SM_State < 100 AND #State > 20 THEN

       //  //     "Control_DB".WMS_OPC_UA.SM_State_Maestro := 3;//RUNNING condition => Shuttle

       //  //     // Any Shuttle Interlock  DONE on the system (Shuttle) 
       //  // ELSIF "Control_DB".WMS_OPC_UA.Task_Type = 2 OR "Control_DB".WMS_OPC_UA.Task_Type = 3
       //  //     AND "Control_DB".WMS_OPC_UA.SM_State = 100 AND #State > 20 THEN

       //  //     "Control_DB".WMS_OPC_UA.SM_State_Maestro := 4;//DONE condition => Shuttle

       //  //     // Any Shuttle Interlock ERRORS on the system (Shuttle) 
       //  // ELSIF "Control_DB".WMS_OPC_UA.Task_Type = 2 OR "Control_DB".WMS_OPC_UA.Task_Type = 3
       //  //     AND "Control_DB".WMS_OPC_UA.SM_State = 400 THEN

       //  //     "Control_DB".WMS_OPC_UA.SM_State_Maestro := 5;//ERROR condition => Shuttle          

       //  // END_IF;

   END_REGION

   #HMI_Reset := ("Screen_DB_1".Reset_All[1] AND
   (("HMI_Box_Connected_1" = 11 AND "KEY REMOTE/LOCAL L1 - CH1(1)") OR
   ("HMI_Box_Connected_1" = 12 AND "KEY REMOTE/LOCAL L2 - CH1(1)") OR
   ("HMI_Box_Connected_1" = 13 AND "KEY REMOTE/LOCAL L3 - CH1(1)") OR
   ("HMI_Box_Connected_1" = 14 AND "KEY REMOTE/LOCAL L4 - CH1(1)") OR
   ("HMI_Box_Connected_1" = 15 AND "KEY REMOTE/LOCAL L5 - CH1(1)") OR
   ("HMI_Box_Connected_1" = 16 AND "KEY REMOTE/LOCAL L6 - CH1(1)") OR
   ("HMI_Box_Connected_1" = 17 AND "KEY REMOTE/LOCAL L7 - CH1(1)") OR
   ("HMI_Box_Connected_1" = 18 AND "KEY REMOTE/LOCAL L8 - CH1(1)") OR
   ("HMI_Box_Connected_1" = 21 AND "KEY REMOTE/LOCAL L1 - CH1(2)") OR
   ("HMI_Box_Connected_1" = 22 AND "KEY REMOTE/LOCAL L2 - CH1(2)") OR
   ("HMI_Box_Connected_1" = 23 AND "KEY REMOTE/LOCAL L3 - CH1(2)") OR
   ("HMI_Box_Connected_1" = 24 AND "KEY REMOTE/LOCAL L4 - CH1(2)") OR
   ("HMI_Box_Connected_1" = 25 AND "KEY REMOTE/LOCAL L5 - CH1(2)") OR
   ("HMI_Box_Connected_1" = 26 AND "KEY REMOTE/LOCAL L6 - CH1(2)") OR
   ("HMI_Box_Connected_1" = 27 AND "KEY REMOTE/LOCAL L7 - CH1(2)") OR
   ("HMI_Box_Connected_1" = 28 AND "KEY REMOTE/LOCAL L8 - CH1(2)") OR
   ("HMI_Box_Connected_1" = 31 AND "KEY REMOTE/LOCAL L1 - CH1(3)") OR
   ("HMI_Box_Connected_1" = 32 AND "KEY REMOTE/LOCAL L2 - CH1(3)") OR
   ("HMI_Box_Connected_1" = 33 AND "KEY REMOTE/LOCAL L3 - CH1(3)") OR
   ("HMI_Box_Connected_1" = 34 AND "KEY REMOTE/LOCAL L4 - CH1(3)") OR
   ("HMI_Box_Connected_1" = 35 AND "KEY REMOTE/LOCAL L5 - CH1(3)") OR
   ("HMI_Box_Connected_1" = 36 AND "KEY REMOTE/LOCAL L6 - CH1(3)") OR
   ("HMI_Box_Connected_1" = 37 AND "KEY REMOTE/LOCAL L7 - CH1(3)") OR
   ("HMI_Box_Connected_1" = 38 AND "KEY REMOTE/LOCAL L8 - CH1(3)") OR
   ("HMI_Box_Connected_1" = 41 AND "KEY REMOTE/LOCAL L1 - CH1(4)") OR
   ("HMI_Box_Connected_1" = 42 AND "KEY REMOTE/LOCAL L2 - CH1(4)") OR
   ("HMI_Box_Connected_1" = 43 AND "KEY REMOTE/LOCAL L3 - CH1(4)") OR
   ("HMI_Box_Connected_1" = 44 AND "KEY REMOTE/LOCAL L4 - CH1(4)") OR
   ("HMI_Box_Connected_1" = 45 AND "KEY REMOTE/LOCAL L5 - CH1(4)") OR
   ("HMI_Box_Connected_1" = 46 AND "KEY REMOTE/LOCAL L6 - CH1(4)") OR
   ("HMI_Box_Connected_1" = 47 AND "KEY REMOTE/LOCAL L7 - CH1(4)") OR
   ("HMI_Box_Connected_1" = 48 AND "KEY REMOTE/LOCAL L8 - CH1(4)") OR
   ("HMI_Box_Connected_1" = 51 AND "KEY REMOTE/LOCAL L1 - CH1(5)") OR
   ("HMI_Box_Connected_1" = 52 AND "KEY REMOTE/LOCAL L2 - CH1(5)") OR
   ("HMI_Box_Connected_1" = 53 AND "KEY REMOTE/LOCAL L3 - CH1(5)") OR
   ("HMI_Box_Connected_1" = 54 AND "KEY REMOTE/LOCAL L4 - CH1(5)") OR
   ("HMI_Box_Connected_1" = 55 AND "KEY REMOTE/LOCAL L5 - CH1(5)") OR
   ("HMI_Box_Connected_1" = 56 AND "KEY REMOTE/LOCAL L6 - CH1(5)") OR
   ("HMI_Box_Connected_1" = 57 AND "KEY REMOTE/LOCAL L7 - CH1(5)") OR
   ("HMI_Box_Connected_1" = 58 AND "KEY REMOTE/LOCAL L8 - CH1(5)")));
END_FUNCTION_BLOCK

FUNCTION_BLOCK "Shuttle_TCP_Comms"   // FB22, SCL
{ S7_Optimized_Access := 'TRUE' }
VERSION : 0.1
// stored: AutoNumber true, IsIECCheckEnabled false, IsRetainMemResEnabled false, MemoryReserve 100, SetENOAutomatically false, UDAEnableTagReadback false
   VAR_INPUT
      Enable : Bool;
      "E-stop" : Bool;
      TCP_Configuration : "LCom_typeConfig";
      Shuttle_No : UInt;
   END_VAR
   VAR_OUTPUT
      Connected : Bool;
      Busy : Bool;
      Status : Word;
      Error : Bool;
   END_VAR
   VAR_IN_OUT
      TCP_Diag : "LCom_typeDiagnostics";
      LCom_Communication_DB : "LCom_Communication_FB";
   END_VAR
   VAR
      SendBuffer { ExternalAccessible := 'False'; ExternalVisible := 'False'; ExternalWritable := 'False'} : Array[0..6] of Byte;
      ReceiveBuffer { ExternalAccessible := 'False'; ExternalVisible := 'False'; ExternalWritable := 'False'} : Array[0..1] of Byte;
      Send : Bool;
      SendDataLength : USInt := 2;
      Sending : Bool;
      T_Send_DB { S7_SetPoint := 'True'} : TON_TIME;
   END_VAR
BEGIN
   IF NOT #"E-stop" THEN
       #SendBuffer[0] := 83;
       IF NOT #Send THEN
           #Send := TRUE;
       END_IF;
   ELSE
       #SendBuffer[0] := 0;
   END_IF;

   #LCom_Communication_DB(enable:=#Enable,
                           send:=#Send,
                           sendDataLength:=#SendDataLength,
                           readDataLength:=16#FFFF_FFFF,
                           configuration:=#TCP_Configuration,
                           connected=>#Connected,
                           sending=>#Sending,
                           busy=>#Busy,
                           error=>#Error,
                           status=>#Status,
                           sendBuffer:=#SendBuffer,
                           receiveBuffer:=#ReceiveBuffer,
                           diagnostics:=#TCP_Diag);


    #SendBuffer[1] := UINT_TO_BYTE("Control_DB".VTD_Sys[1].Current_Level);
    #SendBuffer[2] := UINT_TO_BYTE("Control_DB".VTD_Sys[2].Current_Level);
    #SendBuffer[3] := UINT_TO_BYTE("Control_DB".VTD_Sys[3].Current_Level);
    #SendBuffer[4] := UINT_TO_BYTE("Control_DB".VTD_Sys[4].Current_Level);
    #SendBuffer[5] := UINT_TO_BYTE("Control_DB".VTD_Sys[5].Current_Level);

   "Control_DB".Shuttles_Position[#Shuttle_No].Charging := "Shuttle_MQTT_DB".Shuttle_MQTT[#Shuttle_No].Message.Shuttle_Status.Paused;

   IF #Send AND NOT #Sending THEN
       #Send := FALSE;
   END_IF;

   IF NOT #Send THEN
       #T_Send_DB(IN:=TRUE,
                  PT:=T#500ms);
   END_IF;

   IF #T_Send_DB.Q THEN
       #Send := TRUE;
       #T_Send_DB.TON(IN := FALSE,
                               PT := T#0ms);
   END_IF;
END_FUNCTION_BLOCK

FUNCTION_BLOCK "LCom_Communication_FB"   // FB30300, SCL
TITLE = LCom_Communication
{ S7_Optimized_Access := 'TRUE' }
AUTHOR : APC_ERLF
FAMILY : LCom
VERSION : 2.1
// Support: profinet.team.motioncontrol.i-dt@siemens.com
// Fax: +49 (0) 9131/98-1297
// stored: AutoNumber true, IsIECCheckEnabled false, IsRetainMemResEnabled false, MemoryReserve 100, SetENOAutomatically false, UDAEnableTagReadback false
   VAR_INPUT
      enable : Bool := FALSE;   // Starts the FB with a rising edge
      send : Bool := FALSE;   // Send data connected to input parameter sendBuffer
      sendDataLength : UDInt := 16#FFFF_FFFF;   // Length of data to be sent in Bytes
      readDataLength : UDInt := 16#FFFF_FFFF;   // Receving property: 0 = data from TCP buffer is not read, > 0 = see documentation
      configuration : "LCom_typeConfig";   // FB configuration
   END_VAR
   VAR_OUTPUT
      connected : Bool := FALSE;   // Connection to partner is established
      sending : Bool := FALSE;   // Send data connected to input parameter sendBuffer
      dataReceived : Bool := FALSE;   // New data received
      receivedDataLength : UDInt;   // Length of received data in Bytes
      busy : Bool;   // Processing is executed automatically
      error : Bool := FALSE;   // An error occured
      status : Word := 16#7000;   // FB status
   END_VAR
   VAR_IN_OUT
      sendBuffer : Variant;   // Data to be sent (Array of Byte)
      receiveBuffer : Variant;   // Data received (Array of Byte)
      diagnostics : "LCom_typeDiagnostics";   // Diagnostics
   END_VAR
   VAR
      statConnectAttempts : SInt;
      statActualLocalLComVersion : USInt;
      statRuntimeTask : LReal;
      statCopyNBytes : UDInt;
      statMaxActPacketLength : UDInt;
      statState : Struct
         connection : USInt := 0;
         cfgSender : USInt;
         comSender : USInt;
         comReceiver : USInt;
         sender : USInt;
         receiver : USInt;
      END_STRUCT;
      statReceive : Struct
         tempTelegram : Struct
            LComVersion : USInt;
            index : USInt;
            telegramType : USInt;
            data : Array[0..23] of Byte;
         END_STRUCT;
         configTelegramV1 : Struct
            LComVersion : USInt;
            telegramType : USInt;
            comMode : USInt;
            slidingWindow : USInt;
            cycleTime : UInt;
            ackTimeOut : UInt;
            lifeSignCycle : UInt;
            status : USInt;
            sendModeSyncTime : USInt;
            maxSendDataLength : UInt;
            maxReceiveDataLength : UInt;
         END_STRUCT;
         configTelegramV2 : Struct
            LComVersion : USInt;
            telegramType : USInt;
            status : USInt;
            sendModeSyncTime : USInt;
            lifeSignCycle : Time;
            cycleTime : Time;
            ackTimeOut : Time;
            maxSendDataLength : UDInt;
            maxReceiveDataLength : UDInt;
         END_STRUCT;
         dataTelegram : Struct
            LComVersion : USInt;
            telegramType : USInt;
            messageCounter : USInt;
            ackMessageCounter : USInt;
            messageOffset : UDInt;
            ackMessageOffset : UDInt;
            actPackageLength : UDInt;
            totalMessageLength : UDInt;
         END_STRUCT;
         userData : Struct
            totalLength : UDInt;
            offset : UDInt;
         END_STRUCT;
         trcvFct : Struct
            data : Array[0..4095] of Byte;
            dataOffset : UDInt;
            dataLength : UDInt;
            dataLengthRest : UDInt;
            dataReceived : Bool := FALSE;
         END_STRUCT;
         numberOfLComHeader : USInt;
      END_STRUCT;
      statSend : Struct
         configTelegramV1 : Struct
            LComVersion : USInt;
            comMode : USInt;
            slidingWindow : USInt;
            cycleTime : UInt;
            ackTimeOut : UInt;
            lifeSignCycle : UInt;
            status : USInt;
            sendModeSyncTime : USInt;
            maxSendDataLength : UInt;
            maxReceiveDataLength : UInt;
         END_STRUCT;
         configTelegramV2 : Struct
            LComVersion : USInt;
            status : USInt;
            sendModeSyncTime : USInt;
            lifeSignCycle : Time;
            cycleTime : Time;
            ackTimeOut : Time;
            maxSendDataLength : UDInt;
            maxReceiveDataLength : UDInt;
         END_STRUCT;
         dataTelegram : Struct
            LComVersion : USInt;
            telegramType : USInt;
            messageCounter : USInt;
            ackMessageCounter : USInt;
            messageOffset : UDInt;
            ackMessageOffset : UDInt;
            actPackageLength : UDInt;
            totalMessageLength : UDInt;
         END_STRUCT;
         userData : Struct
            totalLength : UDInt;
            offset : UDInt;
            sendCycleViolation : Bool;
         END_STRUCT;
         tsendFct : Struct
            dataLengthRest : UInt;
            data : Array[0..4095] of Byte;
            dataOffset : UInt;
            status : Word;
            enable : Bool := FALSE;
         END_STRUCT;
         expectedAck : Struct
            package1 : Struct
               offset : UDInt;
            END_STRUCT;
         END_STRUCT;
         numberOfLComPackage : USInt;
      END_STRUCT;
      statIterator : Int;
      statOldEnable : Bool := FALSE;
      statOldSend : Bool := FALSE;
      statRisingEdgeSend : Bool;
      statFallingEdgeEnable : Bool;
      statRet : Int := -1;
      statCompare : Struct
         sender : Struct
            cycleTime : Time;
            ackTimeOut : Time;
         END_STRUCT;
      END_STRUCT;
      statTconPar { S7_SetPoint := 'True'} : TCON_IP_v4;
      statTconParQdn { S7_SetPoint := 'True'} : TCON_QDN;
      instTCON { S7_SetPoint := 'True'} : TCON;
      instTDISCON { S7_SetPoint := 'True'} : TDISCON;
      instTRCV { S7_SetPoint := 'True'} : TRCV;
      instTSEND { S7_SetPoint := 'True'} : TSEND;
      instLocalLifeSignCycleTimer { S7_SetPoint := 'True'} : TON_TIME;
      instPartnerLifeSignCycleTimer { S7_SetPoint := 'True'} : TON_TIME;
      instLocalCycleTimeTimer { S7_SetPoint := 'True'} : TON_TIME;
      instReceiveMsgCycle { S7_SetPoint := 'True'} : TON_TIME;
      instExpectedAckPackage1 { S7_SetPoint := 'True'} : TON_TIME;
      instMsgSendingTimer { S7_SetPoint := 'True'} : TON_TIME;
      instMsgReceivingTimer { S7_SetPoint := 'True'} : TON_TIME;
      instSyncTimer { S7_SetPoint := 'True'} : TON_TIME;
      instSendErrorTimer { S7_SetPoint := 'True'} : TON_TIME;
      instRcvErrorTimer { S7_SetPoint := 'True'} : TON_TIME;
      instRDREC { S7_SetPoint := 'True'} : RDREC;
      statDiag : Struct
         buffer : Array[0..9] of Struct
            status : Word;
            isActive : Bool;
            subFunctionErrorID : Word;
            additionalValue1 : Real;
            additionalValue2 : Real;
            additionalValue3 : Real;
            additionalValue4 : Time;
         END_STRUCT;
         bufferIndex : Int := -1;
         actualIndex : USInt;
      END_STRUCT;
      statDataReceived : Bool;
      statConnected : Bool;
      statStatus : Word;
      statSending : Bool;
   END_VAR
   VAR_TEMP
      tempRuntime : Real;
      tempActTime : DTL;
      tempUDint : UDInt;
      tempDWord : DWord;
      tempConnOucId : CONN_OUC;
   END_VAR
   VAR CONSTANT
      LIFE_SIGN_FACTOR : UInt := 4;
      DIAG_BUFFER_UPPER_LIM : SInt := 63;
      MAX_DATA_BUFFER : Word := 4096;
      HEADER_V1 : USInt := 16#10;
      HEADER_V2 : USInt := 16#20;
      MAX_TRIAL_TIME : Time := T#200MS;
      CON_TYPE_IPV4 : USInt := 1;
      CON_TYPE_QDN : USInt := 10;
      STATE_INACTIVE : USInt;
      STATE_INACTIVE_PREPARE : USInt := 1;
      STATE_INIT : USInt := 2;
      OPEN_SERVER : USInt := 3;
      OPEN_CLIENT : USInt := 4;
      OPERATION : USInt := 5;
      FINISH_TSEND : USInt := 6;
      FINISH_TRCV : USInt := 7;
      CALL_TDISCON : USInt := 8;
      CLOSE_CONNECTION : USInt := 9;
      SEND_CONFIG : USInt := 20;
      SEND_DATA : USInt := 30;
      CYCLE : USInt := 31;
      SEND_NO_DATA : USInt := 38;
      NO_CALL_TRCV : USInt := 40;
      READ : USInt := 50;
      NO_DATA_RECEIVED : USInt := 51;
      DATA_RECEIVED : USInt := 52;
      EXPECTED : USInt := 53;
      DATA_EXPECTED : USInt := 54;
      WAIT_ACK_TELEGRAM : USInt := 55;
      ACK_TELEGRAM : USInt := 56;
      STATE_WAIT : USInt := 60;
      ERROR_STATE : USInt := 99;
      WARN_RECEIVE_BUFFER_LEN : Word := 16#7614;
      ERR_LIFE_SIGN_CYCLE : Word := 16#8210;
      ERR_OPEN_SERVER : Word := 16#8601;
      STATUS_CONNECTED_V1 : Word := 16#7006;
      ERR_COM_SERVICE : Word := 16#8200;
      ERR_ACK_TIMEOUT : Word := 16#8212;
      STATUS_NO_CALL : Word := 16#7000;
      WARN_ACK_TIMEOUT_LIMITATION : Word := 16#7612;
      ERR_WRONG_HEADER : Word := 16#8613;
      ERR_TIME_SYNC_MODE : Word := 16#8205;
      WARN_SEND_CYCLE_EXPIRED : Word := 16#7613;
      STATUS_FIRST_CALL : Word := 16#7001;
      ERR_PARTNER_IP : Word := 16#8204;
      ERR_ACK_MESSAGE_NUMBER : Word := 16#8612;
      ERR_WRONG_TELEGRAM_ID : Word := 16#8614;
      ERR_CONNECTION_ID : Word := 16#8201;
      STATUS_TCP_CONNECTED : Word := 16#7005;
      WARN_LIFE_SIGN_LIMITATION : Word := 16#7610;
      ERR_ACK_TIMEOUT_EXPIRED : Word := 16#8611;
      ERR_SEND_DATA_TYPE : Word := 16#8208;
      ERR_INTERFACE_ID : Word := 16#8202;
      WARN_NO_TIME_SYNC : Word := 16#7615;
      ERR_RECEIVE : Word := 16#8603;
      STATUS_DISCONNECTING : Word := 16#7008;
      STATUS_CLIENT_TRY_CONNECT : Word := 16#7003;
      STATUS_CONNECTED_V2 : Word := 16#7007;
      ERR_RECEIVE_DATA_TYPE : Word := 16#8209;
      ERR_OPEN_CLIENT : Word := 16#8600;
      ERR_LOCAL_PORT : Word := 16#8203;
      ERR_TIME_CYCLE_TIME : Word := 16#8206;
      WARN_SEND_DATA_LENGTH : Word := 16#7600;
      WARN_SEND_CYCLE_LIMITATION : Word := 16#7611;
      ERR_SEND_CYCLE_TIME : Word := 16#8211;
      STATUS_INTERMEDIATE_CALL : Word := 16#7002;
      ERR_SEND : Word := 16#8602;
      ERR_TIME_OF_DAY : Word := 16#8207;
      STATUS_SERVER_PORT_OPEN : Word := 16#7004;
      ERR_LIFE_SIGN_EXPIRED : Word := 16#8610;
      ERR_CLOSE_CONNECTION : Word := 16#8604;
      ERR_CONNECTION_TYPE : Word := 16#8213;
   END_VAR
   // statDiag.buffer[0..9].isActive := FALSE;
BEGIN
   REGION BLOCK INFO HEADER
       //=============================================================================
       // SIEMENS AG / (c)Copyright 2020
       //-----------------------------------------------------------------------------
       // Title:        LCom_Communication
       // Function:     Function block for TCP communication via Industrial Ethernet.
       //               An extended transport protocol, the LCom protocol, has been
       //               implemented for extended communication functions.
       // Library:      LCom
       // Author:       APC_ERLF
       // Tested with:  CPU 1215 V4.x, CPU 1516 V2x
       // Engineering:  TIA Portal V16
       // Restrictions: --
       // Requirements: --
       //-----------------------------------------------------------------------------
       // Change log table:
       // Version  | Date       | Expert in charge       | Changes applied
       //----------|------------|------------------------|------------------------------
       // 02.00.03 | 2015-06-15 | APC_ERLF               | First release
       // 02.00.04 | 2015-09-08 | APC_ERLF               | Several bug fixes
       //                                                | Number of sign-of-life cycles changed from 3 to 4
       // 02.00.05 | 2016-10-10 | APC_ERLF               | Several bug fixes
       //                                                | HW_ANY data type changed (basic data type = UINT)
       // 02.00.06 | 2019-11-07 | APC_ERLF               | Fixed compilation warnings
       // 02.00.07 | 2020.12.16 | APC_ERLF               | Integrated global constants into FB
       // 02.00.08 | 2022.12.01 | APC_ERLF               | Add REGION keywords
       // 02.01.00 | 2022.12.19 | APC_ERLF               | Add connection type (IPv4/QDN) selector in configuration structure
       //=============================================================================
   END_REGION BLOCK INFO HEADER

   REGION RECEIVED_DATA?
       //---------------------------------------------------------------------
       //Reset FB outputs, if in the previous cycle are data received
       //---------------------------------------------------------------------
       IF (#statDataReceived = TRUE) THEN
           #dataReceived := #statDataReceived := FALSE;
           #receivedDataLength := 0;

           //Without LCom protocol
           //Leave the FB, if the tcp buffer is not completely analyzed yet
           //Necessary to enforce an L/H edge (FB.dataReceived), if readDataLength is small
           //Example: Rx=100, readDataLength=1
           IF ((NOT #diagnostics.localConfig.connection.useLComProtocol) AND (#statReceive.trcvFct.dataLengthRest > 0)) THEN
               RETURN;
           END_IF;
       END_IF;
       //End:Reset FB outputs, if in the previous cycle data was received
   END_REGION RECEIVED_DATA?

   REGION ENABLING/DISABLING
       //---------------------------------------------------------------------
       //Check enable input
       //---------------------------------------------------------------------
       IF ((#enable) AND (NOT #statOldEnable) AND (NOT #statFallingEdgeEnable))//Rising edge
       THEN
           //Start initialize state for the tcp connection
           #statState.connection := #STATE_INIT;
           #status := #statStatus := #STATUS_FIRST_CALL;
           #busy := TRUE;
       ELSIF (NOT #enable AND #statState.connection = #STATE_INACTIVE) THEN//Inactive
           RETURN;//Do nothing, wait rising edge on enable
       ELSIF ((NOT #enable) AND (#statOldEnable)) THEN//Falling edge

           #statFallingEdgeEnable := TRUE;
           //LCom Version 1.0 or 2.0 is used OR native tcp
           #statState.connection := #CLOSE_CONNECTION;

           #status := #statStatus := #STATUS_DISCONNECTING;
           //Write diagnostics
           #statDiag.bufferIndex := #statDiag.bufferIndex + 1;
           #statDiag.buffer[#statDiag.bufferIndex].status := #STATUS_DISCONNECTING;
           #statDiag.buffer[#statDiag.bufferIndex].subFunctionErrorID := 16#0000;
           #statDiag.buffer[#statDiag.bufferIndex].additionalValue1 := 0.0;
           #statDiag.buffer[#statDiag.bufferIndex].additionalValue2 := 0.0;
           #statDiag.buffer[#statDiag.bufferIndex].additionalValue3 := 0.0;
           #statDiag.buffer[#statDiag.bufferIndex].additionalValue4 := T#0ms;
       ELSE
           ;//No change on enable input
       END_IF;
       #statOldEnable := #enable;
       //End:Check enable input
   END_REGION ENABLING/DISABLING

   REGION CYCLE_TIME_STATISTIC
       // -----------------------------------------------------------------------------------------------------------
       //Statistic --> Calculate average of cycle time [ms]
       // -----------------------------------------------------------------------------------------------------------
       #tempRuntime := (LREAL_TO_REAL(RUNTIME(#statRuntimeTask)) * 1000);

       //Check the measured runtime value and calculate average of cycle time
       IF ((#tempRuntime > 0) AND #enable)
       THEN
           #diagnostics.statistics.avgCallCycle := (((#diagnostics.statistics.avgCallCycle * 49.0) + #tempRuntime) / 50.0);
       ELSE
           ;//Ignore this runtime value 
       END_IF;
   END_REGION CYCLE_TIME_STATISTIC

   REGION INIT_VALUES
       //---------------------------------------------------------------------
       //Initialize values
       //---------------------------------------------------------------------
       #statState.sender := #STATE_INACTIVE;
       #statSend.tsendFct.enable := FALSE;
       #statSend.tsendFct.dataOffset := 0;
       //Set index of temp diagnostics entry
       #statDiag.bufferIndex := -1;
       //End: Calculate average of cycle time and initialize values
   END_REGION INIT_VALUES

   REGION CHECK_SEND_INPUT
       //---------------------------------------------------------------------
       //Check send input
       //---------------------------------------------------------------------
       IF #statConnected THEN
           //Check rising edge
           IF (#send AND (NOT #statOldSend)) THEN
               //Rising edge detected
               #statRisingEdgeSend := TRUE;
           ELSE
               ;
           END_IF;
           #statOldSend := #send;
       ELSE
           ;//Change at send input is not relevant, because FB is not connected
       END_IF;
       //End:Check send input
   END_REGION CHECK_SEND_INPUT

   REGION ACK_AUTOMATICALLY_WARNINGS
       //---------------------------------------------------------------------
       //Acknowledge automatically the followings warnings
       //---------------------------------------------------------------------
       IF (#statStatus = #WARN_SEND_DATA_LENGTH)
           OR (#statStatus = #WARN_SEND_CYCLE_EXPIRED)
           OR (#statStatus = #WARN_RECEIVE_BUFFER_LEN
           OR (#statStatus = #WARN_NO_TIME_SYNC))
       THEN
           //With LCom protocol
           IF #diagnostics.localConfig.connection.useLComProtocol THEN

               IF (#diagnostics.statistics.activeLComVersion = #HEADER_V1) THEN
                   #status := #STATUS_CONNECTED_V1;
               ELSE
                   #status := #STATUS_CONNECTED_V2;
               END_IF;
           ELSE//Without LCom protocol
               #status := #statStatus := #STATUS_TCP_CONNECTED;
           END_IF;
       END_IF;
       //End:Acknowledge automatically the followings warnings
   END_REGION ACK_AUTOMATICALLY_WARNINGS

   REGION STATE_MACHINE
       //---------------------------------------------------------------------
       // State machine for IP connection
       //---------------------------------------------------------------------
       CASE #statState.connection OF

           #OPERATION:
               REGION OPERATION
                   //IP connection is established

                   REGION CHECK_LIFESIGN
                       //Get time difference between the last received telegram
                       #instPartnerLifeSignCycleTimer(IN := TRUE,
                                                      PT := (#diagnostics.partnerConfig.connnection.lifeSignCycleTime * #LIFE_SIGN_FACTOR));

                       //Only with LCom protocol, check life sign monitoring
                       IF ((#diagnostics.localConfig.connection.useLComProtocol)
                           AND
                           (#diagnostics.partnerConfig.connnection.lifeSignCycleTime > T#0ms)
                           AND
                           (#instPartnerLifeSignCycleTimer.Q))
                       THEN
                           //Write diagnostics
                           #statDiag.bufferIndex := #statDiag.bufferIndex + 1;
                           #statDiag.buffer[#statDiag.bufferIndex].status := #ERR_LIFE_SIGN_EXPIRED;
                           #statDiag.buffer[#statDiag.bufferIndex].subFunctionErrorID := 16#0000;
                           #statDiag.buffer[#statDiag.bufferIndex].additionalValue1 := UDINT_TO_REAL(TIME_TO_UDINT(#diagnostics.partnerConfig.connnection.lifeSignCycleTime));
                           #statDiag.buffer[#statDiag.bufferIndex].additionalValue2 := 0.0;
                           #statDiag.buffer[#statDiag.bufferIndex].additionalValue3 := 0.0;
                           #statDiag.buffer[#statDiag.bufferIndex].additionalValue4 := #instPartnerLifeSignCycleTimer.ET;

                           #statState.connection := #CLOSE_CONNECTION;
                           GOTO diag;
                       END_IF;
                   END_REGION CHECK_LIFESIGN

                   REGION CHECK_SENDING
                       //---------------------------------------------------------------------
                       //Check the status of the "TSEND" instruction of the previous request
                       //---------------------------------------------------------------------
                       IF ((#statSend.tsendFct.status = 16#7001)
                           OR
                           (#statSend.tsendFct.status = 16#7002)
                           OR
                           (#statSend.tsendFct.status = 16#80C4))
                       THEN
                           //differ between different connection types (IPv4, QDN)
                           IF (#diagnostics.localConfig.connection.connectType = #CON_TYPE_IPV4) THEN
                               #tempConnOucId := #statTconPar.ID;
                           ELSE    //#CON_TYPE_QDN
                               #tempConnOucId := #statTconParQdn.ID;
                           END_IF;
                           //When "TSEND" instruction started or is in sending process
                           #instTSEND(REQ := TRUE,
                                      LEN := #statSend.tsendFct.dataOffset,
                                      ID := #tempConnOucId,
                                      DATA := #statSend.tsendFct.data,
                                      STATUS => #statSend.tsendFct.status);

                           //When "TSEND" instruction of the previous request is not yet completed
                           IF ((#statSend.tsendFct.status = 16#7001)
                               OR
                               (#statSend.tsendFct.status = 16#7002))
                           THEN
                               //Stop SendError timer
                               #instSendErrorTimer(IN := FALSE,
                                                   PT := #MAX_TRIAL_TIME);
                               RETURN;//"TSEND" instruction still in process, leave FB
                           ELSIF (#statSend.tsendFct.status = 16#80C4) THEN
                               //Temporary communication error-->Start/Get SendError timer
                               #instSendErrorTimer(IN := TRUE,
                                                   PT := #MAX_TRIAL_TIME);

                               //#MAX_TRIAL_TIME is expired
                               IF #instSendErrorTimer.Q THEN
                                   //Write diagnostics
                                   #statDiag.bufferIndex := #statDiag.bufferIndex + 1;
                                   #statDiag.buffer[#statDiag.bufferIndex].status := #ERR_SEND;
                                   #statDiag.buffer[#statDiag.bufferIndex].subFunctionErrorID := #statSend.tsendFct.status;
                                   #statDiag.buffer[#statDiag.bufferIndex].additionalValue1 := 0.0;
                                   #statDiag.buffer[#statDiag.bufferIndex].additionalValue2 := #statSend.tsendFct.dataOffset;
                                   #statDiag.buffer[#statDiag.bufferIndex].additionalValue3 := 0.0;
                                   #statDiag.buffer[#statDiag.bufferIndex].additionalValue4 := T#0ms;
                                   #statState.connection := #CLOSE_CONNECTION;
                                   GOTO diag;
                               ELSE
                                   RETURN;//Temporary communication error still valid ant timer is not expired leave FB
                               END_IF;
                           ELSIF ((#statSend.tsendFct.status = 16#7000) OR (#statSend.tsendFct.status = 16#0000)) THEN
                               //---------------------------------------------------------------------
                               //Send job completed without error
                               //---------------------------------------------------------------------
                               IF ((NOT #diagnostics.localConfig.connection.useLComProtocol)
                                   AND
                                   (#statSend.userData.offset = #statSend.dataTelegram.totalMessageLength))
                               THEN
                                   //Without LCom protocol
                                   #statSend.dataTelegram.totalMessageLength := 0;
                                   #sending := #statSending := FALSE;

                                   //Statistic, increase number of sent messages
                                   #diagnostics.statistics.numberOfSentMessages := #diagnostics.statistics.numberOfSentMessages + 1;

                                   //Get the message sending time (ms)
                                   #instMsgSendingTimer(IN := TRUE,
                                                        PT := T#+24d20h31m23s647ms);

                                   //Check maximum message sending time (ms)
                                   IF (#instMsgSendingTimer.ET > #diagnostics.statistics.maxMsgSendingTime) THEN
                                       #diagnostics.statistics.maxMsgSendingTime := #instMsgSendingTimer.ET;
                                   ELSE
                                       ;//Actual sending time is smaller
                                   END_IF;

                                   //Calculate average of message sending time (ms)
                                   #diagnostics.statistics.avgMsgSendingTime := (((#diagnostics.statistics.avgMsgSendingTime * 19) + UDINT_TO_REAL((TIME_TO_UDINT(#instMsgSendingTimer.ET)))) / 20);

                                   //Stop message sending timer
                                   #instMsgSendingTimer(IN := FALSE,
                                                        PT := T#+24d20h31m23s647ms);
                               ELSE
                                   ;//With LCom protocol and not in disconnecting process
                               END_IF;
                               //Stop SendError timer
                               #instSendErrorTimer(IN := FALSE,
                                                   PT := #MAX_TRIAL_TIME);

                               //Call "TSEND" instruction, with REQ:= FALSE (falling edge)
                               //Preparation for the next send job
                               #instTSEND(REQ := FALSE,
                                          LEN := #statSend.tsendFct.dataOffset,
                                          ID := #tempConnOucId,
                                          DATA := #statSend.tsendFct.data,
                                          STATUS => #statSend.tsendFct.status);

                               #statSend.tsendFct.dataOffset := 0;
                               //End:Send job completed without error
                           ELSE
                               //An error occurred during execution of "TSEND" call
                               //The data to send was not completely transmitted
                               //Write diagnostics
                               #statDiag.bufferIndex := #statDiag.bufferIndex + 1;
                               #statDiag.buffer[#statDiag.bufferIndex].status := #ERR_SEND;
                               #statDiag.buffer[#statDiag.bufferIndex].subFunctionErrorID := #statSend.tsendFct.status;
                               #statDiag.buffer[#statDiag.bufferIndex].additionalValue1 := 0.0;
                               #statDiag.buffer[#statDiag.bufferIndex].additionalValue2 := #statSend.tsendFct.dataOffset;
                               #statDiag.buffer[#statDiag.bufferIndex].additionalValue3 := 0.0;
                               #statDiag.buffer[#statDiag.bufferIndex].additionalValue4 := T#0ms;

                               #statState.connection := #CLOSE_CONNECTION;
                               GOTO diag;
                           END_IF;
                       ELSE
                           ; //The "TSEND" instruction is not started or in processing
                       END_IF;
                       //End:Check the #status OF the TSEND instruction from the previous request
                   END_REGION CHECK_SENDING

                   REGION READ_TCP_BUFFER
                       //Check if the tcp buffer must read
                       IF (#readDataLength = 0 OR #statState.cfgSender = #STATE_INIT OR #statState.cfgSender = #SEND_CONFIG)
                       THEN
                           ;//Do not read tcp Buffer
                       ELSE
                           //Check if there are still data in the tcp buffer from the previous "TRCV" call
                           IF (#statState.receiver = #NO_CALL_TRCV) THEN
                               ;//Still bytes in the tcp buffer, don´t call "TRCV" instruction
                           ELSE
                               //Read the complete tcp buffer
                               #instTRCV.STATUS := 16#0000;
                               #instTRCV(EN_R := TRUE,
                                         ID := #diagnostics.localConfig.connection.connectionID,
                                         LEN := 0,
                                         ADHOC := TRUE,
                                         NDR => #statReceive.trcvFct.dataReceived,
                                         RCVD_LEN => #statReceive.trcvFct.dataLength,
                                         DATA := #statReceive.trcvFct.data);

                               //An error occurred during execution of "TRCV" call
                               IF (#instTRCV.ERROR) THEN
                                   //16#80C4=Temporary communication error
                                   //16#80A1=Connection or port already being used by user
                                   IF ((#instTRCV.STATUS = 16#80C4) OR (#instTRCV.STATUS = 16#80A1)) THEN
                                       //Get RcvError time
                                       #instRcvErrorTimer(IN := TRUE,
                                                          PT := #MAX_TRIAL_TIME);

                                       //#MAX_TRIAL_TIME is expired
                                       IF #instRcvErrorTimer.Q THEN
                                           //Write diagnostics
                                           #statDiag.bufferIndex := #statDiag.bufferIndex + 1;
                                           #statDiag.buffer[#statDiag.bufferIndex].status := #ERR_RECEIVE;
                                           #statDiag.buffer[#statDiag.bufferIndex].subFunctionErrorID := #instTRCV.STATUS;
                                           #statDiag.buffer[#statDiag.bufferIndex].additionalValue1 := 0.0;
                                           #statDiag.buffer[#statDiag.bufferIndex].additionalValue2 := 0.0;
                                           #statDiag.buffer[#statDiag.bufferIndex].additionalValue3 := 0.0;
                                           #statDiag.buffer[#statDiag.bufferIndex].additionalValue4 := T#0ms;
                                           #statState.connection := #CLOSE_CONNECTION;
                                           GOTO diag;
                                       END_IF;
                                       //Stop partner watch dog timer of life sign cycle
                                       #instPartnerLifeSignCycleTimer(IN := FALSE,
                                                                      PT := (#diagnostics.partnerConfig.connnection.lifeSignCycleTime * #LIFE_SIGN_FACTOR));
                                   ELSE//An error occurred during execution <>16#80C4 and <> 16#80A1
                                       //Write diagnostics
                                       #statDiag.bufferIndex := #statDiag.bufferIndex + 1;
                                       #statDiag.buffer[#statDiag.bufferIndex].status := #ERR_RECEIVE;
                                       #statDiag.buffer[#statDiag.bufferIndex].subFunctionErrorID := #instTRCV.STATUS;
                                       #statDiag.buffer[#statDiag.bufferIndex].additionalValue1 := 0.0;
                                       #statDiag.buffer[#statDiag.bufferIndex].additionalValue2 := 0.0;
                                       #statDiag.buffer[#statDiag.bufferIndex].additionalValue3 := 0.0;
                                       #statDiag.buffer[#statDiag.bufferIndex].additionalValue4 := T#0ms;
                                       #statState.connection := #CLOSE_CONNECTION;
                                       GOTO diag;
                                   END_IF;
                               ELSE
                                   //"TRCV" call completed without error
                                   //New data received
                                   IF (#instTRCV.NDR) THEN

                                       #statState.receiver := #DATA_RECEIVED;

                                       //Stop partner watch dog timer of life sign cycle
                                       #instPartnerLifeSignCycleTimer(IN := FALSE,
                                                                      PT := (#diagnostics.partnerConfig.connnection.lifeSignCycleTime * #LIFE_SIGN_FACTOR));

                                       #statReceive.trcvFct.dataLengthRest := #statReceive.trcvFct.dataLength;
                                       #statReceive.trcvFct.dataOffset := 0;

                                       //Reset the counter
                                       #statCopyNBytes := 0;
                                   ELSE
                                       //No data received
                                       #statState.receiver := #NO_DATA_RECEIVED;
                                   END_IF;
                                   //Stop RcvError timer
                                   #instRcvErrorTimer(IN := FALSE,
                                                      PT := #MAX_TRIAL_TIME);
                               END_IF;
                           END_IF;

                           //Initialize before the tcp is analyzed
                           #statReceive.numberOfLComHeader := 0;

                           //---------------------------------------------------------------------
                           //Analysis tcp receive buffer
                           //---------------------------------------------------------------------
                           REPEAT

                               //The complete tcp receive buffer is analyzed --> stop analyzing
                               IF (#statReceive.trcvFct.dataLengthRest <= 0)
                               THEN
                                   EXIT;
                               END_IF;
                               REGION NATIVE_TCP
                                   //---------------------------------------------------------------------
                                   //Analyze tcp receive buffer without LCom protocol
                                   //---------------------------------------------------------------------
                                   IF (NOT #diagnostics.localConfig.connection.useLComProtocol) THEN

                                       //Store the total receive length with the 1st received telegram
                                       IF (#statReceive.userData.offset = 0) THEN

                                           //Compare readDataLength with the local max. receive data length
                                           IF ((#diagnostics.localConfig.sizeOfReceiveBuffer < #readDataLength)
                                               AND
                                               (#readDataLength > 0 AND #readDataLength < 4294967295))//#readDataLength 1 ... 4294967295
                                           THEN
                                               #statDiag.bufferIndex := #statDiag.bufferIndex + 1;
                                               #statDiag.buffer[#statDiag.bufferIndex].status := #WARN_RECEIVE_BUFFER_LEN;
                                               #statDiag.buffer[#statDiag.bufferIndex].subFunctionErrorID := 16#0000;
                                               #statDiag.buffer[#statDiag.bufferIndex].additionalValue1 := UDINT_TO_REAL(#diagnostics.localConfig.sizeOfReceiveBuffer);

                                               #statDiag.buffer[#statDiag.bufferIndex].additionalValue2 := UDINT_TO_REAL(#readDataLength);
                                               #statDiag.buffer[#statDiag.bufferIndex].additionalValue3 := 0.0;
                                               #statDiag.buffer[#statDiag.bufferIndex].additionalValue4 := T#0ms;

                                               #statReceive.userData.totalLength := #diagnostics.localConfig.sizeOfReceiveBuffer;
                                           ELSIF (#readDataLength = 4294967295) THEN//Adhoc
                                               //The TRCV Fkt. can read up to 4096 Byte
                                               //If the Rx user buffer is less than the current received bytes, limit to the Rx user buffer
                                               //Otherwise copy received bytes (LCom internal Rx) to the Rx user buffer
                                               IF (#statReceive.trcvFct.dataLengthRest < #diagnostics.localConfig.sizeOfReceiveBuffer)
                                               THEN
                                                   #statReceive.userData.totalLength := #statReceive.trcvFct.dataLengthRest;
                                               ELSE
                                                   #statReceive.userData.totalLength := #diagnostics.localConfig.sizeOfReceiveBuffer;
                                               END_IF;
                                           ELSE
                                               #statReceive.userData.totalLength := #readDataLength;
                                           END_IF;

                                           //Start message receiving timer (ms)
                                           //Duration between start of message and FB output dataReceived becomes TRUE
                                           #instMsgReceivingTimer(IN := TRUE,
                                                                  PT := T#+24d20h31m23s647ms);
                                       ELSE
                                           ;//Not the 1st received telegram
                                       END_IF;

                                       //Is the data to be analyzed in the tcp receive buffer bigger than the complete message ?
                                       IF (#statReceive.userData.offset + #statReceive.trcvFct.dataLengthRest) > #statReceive.userData.totalLength THEN
                                           //Copy only the rest data from the message, not all data from the tcp receive buffer
                                           #statCopyNBytes := #statReceive.userData.totalLength - #statReceive.userData.offset;
                                       ELSE
                                           //Copy just the rest of data from the tcp receive buffer
                                           #statCopyNBytes := #statReceive.trcvFct.dataLengthRest;
                                       END_IF;

                                       //Copy data to FB.receiveBuffer
                                       #statRet := MOVE_BLK_VARIANT(SRC := #statReceive.trcvFct.data, COUNT := #statCopyNBytes, SRC_INDEX := UDINT_TO_DINT(#statReceive.trcvFct.dataOffset), DEST_INDEX := UDINT_TO_DINT(#statReceive.userData.offset), DEST => #receiveBuffer);
                                       //Calculate offset in the FB.#receiveBuffer
                                       #statReceive.userData.offset := #statReceive.userData.offset + #statCopyNBytes;
                                       //Calculate offset in the tcp receive buffer
                                       #statReceive.trcvFct.dataOffset := #statReceive.trcvFct.dataOffset + #statCopyNBytes;
                                       //Calculate the rest of data in the tcp receive buffer
                                       #statReceive.trcvFct.dataLengthRest := #statReceive.trcvFct.dataLength - #statReceive.trcvFct.dataOffset;

                                       //Is the complete message in the FB.#receiveBuffer copied ?
                                       IF (#statReceive.userData.offset = #statReceive.userData.totalLength) THEN
                                           //The complete message is copied in the FB.#receiveBuffer
                                           //Set FB outputs and initialize for the next receive request
                                           #dataReceived := #statDataReceived := TRUE;
                                           #receivedDataLength := #statReceive.userData.totalLength;
                                           #statReceive.userData.offset := 0;

                                           //Statistic --> increase number of received user messages
                                           #diagnostics.statistics.numberOfReceivedMessages := #diagnostics.statistics.numberOfReceivedMessages + 1;

                                           //Get message receiving time [ms]
                                           #instMsgReceivingTimer(IN := TRUE,
                                                                  PT := T#+24d20h31m23s647ms);

                                           //Statistic --> compare max. message receiving time
                                           IF (#instMsgReceivingTimer.ET > #diagnostics.statistics.maxMsgReceivingTime) THEN
                                               #diagnostics.statistics.maxMsgReceivingTime := #instMsgReceivingTimer.ET;
                                           ELSE
                                               ;//Actual receiving time is smaller
                                           END_IF;

                                           //Statistic --> calculate average of message receiving time (ms)
                                           #diagnostics.statistics.avgMsgReceivingTime := (((#diagnostics.statistics.avgMsgReceivingTime * 19) + UDINT_TO_REAL((TIME_TO_UDINT(#instMsgReceivingTimer.ET)))) / 20);

                                           //Stop message receiving timer
                                           #instMsgReceivingTimer(IN := FALSE,
                                                                  PT := T#+24d20h31m23s647ms);

                                           //Get receive message cycle time [ms]
                                           #instReceiveMsgCycle(IN := TRUE,
                                                                PT := T#+24d20h31m23s647ms);

                                           //Statistic --> compare max. receive message cycle time
                                           IF (#instReceiveMsgCycle.ET > #diagnostics.statistics.maxReceiveMsgCycle) THEN
                                               #diagnostics.statistics.maxReceiveMsgCycle := #instReceiveMsgCycle.ET;
                                           ELSE
                                               ;//Actual receive message cycle time is smaller
                                           END_IF;

                                           //Statistic --> calculate average of receive message cycle time
                                           #diagnostics.statistics.avgReceiveMsgCycle := (((#diagnostics.statistics.avgReceiveMsgCycle * 19) + UDINT_TO_REAL((TIME_TO_UDINT(#instReceiveMsgCycle.ET)))) / 20);

                                           //Stop receive message cycle timer
                                           #instReceiveMsgCycle(IN := FALSE,
                                                                PT := T#+24d20h31m23s647ms);

                                           //Start receive message cycle timer
                                           #instReceiveMsgCycle(IN := TRUE,
                                                                PT := T#+24d20h31m23s647ms);

                                           //There are still bytes in the tcp receive buffer which must be analyzed
                                           IF (#statReceive.trcvFct.dataLengthRest > 0) THEN
                                               //Do not call "TRCV" instruction
                                               #statState.receiver := #NO_CALL_TRCV;
                                           ELSE
                                               //Call "TRCV" instruction in the next cycle
                                               #statState.receiver := #READ;
                                           END_IF;
                                       ELSE
                                           //The complete message is not copied to the FB.#receiveBuffer
                                           #statState.receiver := #READ;
                                       END_IF;
                                       EXIT;//Stop analyzing the tcp receive buffer without LCom protocol
                                   ELSE
                                       ;//With LCom protocol
                                   END_IF;//End: Analyze tcp receive buffer without LCom protocol
                               END_REGION NATIVE_TCP

                               REGION LCOM_PROTOCOL
                                   //---------------------------------------------------------------------
                                   //Analyze tcp receive buffer with LCom protocol
                                   //---------------------------------------------------------------------

                                   //Is data expected without LCom header ?
                                   IF (#statState.comReceiver = #DATA_EXPECTED) THEN
                                       ;//LCom header is already known, still some bytes missing so the actual LCom package becomes complete
                                   ELSE
                                       //There is already data in the temp. LCom header ?
                                       IF (#statReceive.tempTelegram.index = 0) THEN
                                           //No data in the temp. LCom header
                                           //Get the LCom version from the receive telegram
                                           #statReceive.tempTelegram.LComVersion := #statReceive.trcvFct.data[#statReceive.trcvFct.dataOffset];

